(* IEC 61131-3 sources: daoli-st-library/DL_MathData (part 29) *)

(* ---- FB_DL_MovingAverage.st ---- *)
(*==============================================================================
 * 组件名称 (Component)  : FB_DL_MovingAverage
 * 所属子库 (Sublibrary) : DL_MathData
 * 当前版本 (Version)    : 1.0.0
 * 兼容性   (Platform)   : CODESYS 3.5 / TwinCAT 3 / 汇川 InoProShop / Machine Expert
 *                         仅依赖 Standard.library（R_TRIG），全 REAL 运算
 * 功能描述 (Function)   : O(1) 递推滑动平均滤波。窗口长度运行时可改，采样节拍由
 *                         调用方控制。两阶段启动：窗口未满阶段只"写入+累加+计数"、
 *                         绝不执行"减最旧值"；窗口已满阶段执行"减最旧+加最新+指针递增"。
 *                         每 DL_MAV_CORRECT_CYCLE 次采样做一次全窗口重算，消除浮点
 *                         累加漂移。窗口长度变更时整体重建缓冲区，避免新旧样本混算产生台阶。
 *
 * 【滞后披露 / Phase lag disclosure（边界 B11）】
 *   相位滞后约 (N-1)/2 个采样周期，滤波时间窗 = N × 采样周期。
 *   安全联锁回路（急停、超压保护、超温切断）严禁使用大窗口滤波值，
 *   必须直接使用原始信号或小窗口（N ≤ 3）值。
 *
 * 【断电保持提示 / Retain hint（边界 B12）】
 *   缓冲区、写指针、累加和、已填充数若不设 RETAIN，重新上电会重走"窗口未满"阶段，
 *   表现为输出从 0 缓慢爬升。需要无扰重启的场合，应将本实例声明为 VAR RETAIN。
 *
 * 【采样语义 / Sampling semantics（边界 B7，重要）】
 *   采样判据统一为"bSample 电平为 TRUE 即采样"：bSample := TRUE 常 TRUE 时每周期采样，
 *   接一个上升沿脉冲变量则按事件采样。绝不用 R_TRIG 承担两种语义——常 TRUE 信号经
 *   R_TRIG 只在首周期产生一次脉冲，会导致"只采到一个样本"的低级事故。
 *   因此本组件不设 fbTrigSample 采样沿实例（仅保留 fbTrigReset），
 *   这是对 ROUND_PLAN §2.13 VAR 清单的刻意收窄，依据 B7 与决策记录 P6。
 *
 * 【状态机 / State machine（边界 B1/B10）】
 *   采用 eInit / eFilling / eRunning / eFault 四态 + ELSE 兜底。
 *   两阶段判据由 bBufferFull 承担并在采样段用 IF bBufferFull THEN … ELSE … END_IF（代码骨架，示例省略）
 *   显式分支，采样算术只写一处，状态机只负责阶段迁移，避免同一段代码在两个 CASE
 *   分支中重复而导致"只改一处"的缺陷。
 * 开源溯源 (Origin)     : 原创实现。环形缓冲 + 递推求和的滑动平均为公开经典算法。
 * 依赖     (Depends)    : 无 DL_ 内部依赖；Standard.library: R_TRIG
 * 红线自检 (Redline)    : R1 ✓ 零全局变量表与外部变量引用 ｜ R2 ✓ 零物理 IO 地址直写
 *                         R3 ✓ 纯 IEC 61131-3 ｜ R4 ✓ 除零双保险/窗口钳位/MOD 回绕/重算防死锁
 *                         R5 ✓ 全变量中英双语同行注释 ｜ R6 ✓ 四态 ENUM+CASE+ELSE 兜底
 *                         R7 ✓ R_TRIG 主体最前部无条件刷新
 * 修订历史 (Revision)   :
 *   2026-11-14  v1.0.0  首版入库（Phase 1 冷启动 · Level 0 批次）
 *============================================================================*)

(*-----------------------------------------------------------------------------
 * 枚举: E_DL_MovingAverageState（归属 DL_MathData，与 FB_DL_MovingAverage 同文件）
 * 含义: 滑动平均工作阶段。eFilling 与 eRunning 的区分仅用于状态迁移与诊断，
 *       采样算术由 bBufferFull 在单一分支内完成。
 *----------------------------------------------------------------------------*)
TYPE E_DL_MovingAverageState :
(
    eInit    := 0,    // 初始化态：清缓冲、清累加和、清故障，单周期驻留 / Initialization: clear buffer, sum and fault, single scan
    eFilling := 10,   // 填充态：窗口未满，只追加样本不做淘汰 / Filling: window not full, append only without eviction
    eRunning := 20,   // 运行态：窗口已满，执行 O(1) 递推替换 / Running: window full, O(1) recursive replacement
    eFault   := 99    // 故障态：非法状态命中，输出保持最后有效值 / Fault: illegal state hit, outputs hold the last valid value
);
END_TYPE

FUNCTION_BLOCK FB_DL_MovingAverage
VAR_INPUT
    fInput      : REAL := 0.0;      // 原始采样值 [EU] / Raw sampled value [EU]
    nWindowSize : INT := 8;         // 窗口长度，合法域 1..100 / Window length, valid range 1..100
    bSample     : BOOL := TRUE;     // 采样触发，电平 TRUE 即采样；接脉冲变量则按事件采样 / Sample trigger, TRUE level samples every scan
    bEnable     : BOOL := TRUE;     // 使能标志，FALSE 时停止采样并保持输出 / Enable flag, FALSE stops sampling and holds the output
    bReset      : BOOL;             // 复位信号，上升沿清空窗口与累加和 / Reset, rising edge clears the buffer and the sum
END_VAR
VAR_OUTPUT
    fAverage     : REAL;            // 窗口算术平均 [EU] / Window arithmetic mean [EU]
    bBufferFull  : BOOL;            // 窗口已填满标志，同时作为两阶段判据 / Buffer full flag, also the two-phase discriminator
    nSampleCount : INT;             // 窗口内有效样本数，值域 0..nWindowSize / Valid sample count in the window, range 0..nWindowSize
    fWindowSum   : REAL;            // 窗口累加和，诊断用 [EU] / Window sum for diagnostics [EU]
    bError       : BOOL;            // 故障标志，需 bReset 清除 / Fault flag, cleared by bReset
    uErrorId     : UDINT;           // 故障码，0 = 无故障 / Error code, 0 = no error
END_VAR
VAR
    afBuffer     : ARRAY[0..99] OF REAL;  // 环形缓冲区，容量等于窗口上限 [EU] / Ring buffer sized to the max window [EU]
    nWriteIndex  : INT;             // 环形写指针，值域 0..99 / Ring write index, range 0..99
    nFilled      : INT;             // 已填充样本数，值域 0..100 / Number of filled samples, range 0..100
    fSum         : REAL;            // 滑动累加和 [EU]，与 nFilled 同步维护 / Running sum [EU], maintained with nFilled
    nLastWindow  : INT;             // 上周期窗口长度，用于变更检测 / Previous window length for change detection
    fbTrigReset  : R_TRIG;          // 复位上升沿检测实例 / Reset rising edge detector instance
    nCorrectCnt  : DINT;            // 距下次全窗口重算的采样计数 / Sample counter until the next full-window recalculation
    nGuard       : DINT;            // 重算循环防死锁计数器 / Recalculation loop deadlock guard
    fRecalcSum   : REAL;            // 重算中间累加和 [EU] / Recalculation intermediate sum [EU]
    nIdx         : INT;             // 重算循环索引，值域 0..99 / Recalculation loop index, range 0..99
    nWindowEff   : INT;             // 钳位后的有效窗口长度 / Clamped effective window length
    eState       : E_DL_MovingAverageState; // 主状态机当前状态 / Current state of the main state machine
    bDoSample    : BOOL;            // 本周期采样使能（bSample AND bEnable） / Sampling enabled this scan
    bJustReset   : BOOL;            // 本周期刚发生复位/初始化，需跳过采样 / Reset or init happened this scan, sampling is skipped
END_VAR
VAR CONSTANT
    DL_MAV_MAX_WINDOW    : INT := 100;        // 窗口上限，必须与数组维度一致 / Max window, must match the array dimension
    DL_MAV_MIN_WINDOW    : INT := 1;          // 窗口下限 / Min window
    DL_MAV_CORRECT_CYCLE : DINT := 10000;     // 每 N 次采样做一次全窗口重算校正 / Recalculate every N samples
    DL_MAV_MAX_LOOP      : DINT := 100;       // 重算循环迭代上限 / Recalculation loop iteration limit
    DL_FLOAT_EPS         : REAL := 1.0E-6;    // 浮点判零容差 / Float zero tolerance
END_VAR

(*------------------------------------------------------------------------------
 * 段 1｜无条件刷新区（红线 R7）：复位沿实例在主体最前部调用，严禁进入 IF/CASE
 *      Unconditional refresh zone: the reset edge instance runs at the very top
 *-----------------------------------------------------------------------------*)
fbTrigReset(CLK := bReset);

(*------------------------------------------------------------------------------
 * 段 2｜窗口长度钳位（边界 B3）：先钳位，后用于所有后续计算
 *      Window length clamping: clamp first, then use everywhere
 *------------------------------------------------------------------------------*)
IF nWindowSize < DL_MAV_MIN_WINDOW THEN
    nWindowEff := DL_MAV_MIN_WINDOW;
    uErrorId   := 16#0001_0001;
    bError     := TRUE;
ELSIF nWindowSize > DL_MAV_MAX_WINDOW THEN
    nWindowEff := DL_MAV_MAX_WINDOW;
    uErrorId   := 16#0001_0001;
    bError     := TRUE;
ELSE
    nWindowEff := nWindowSize;
END_IF

(*------------------------------------------------------------------------------
 * 段 3｜窗口长度变更重建（边界 B4）：清空缓冲、指针、累加和，重走未满阶段
 *      Window change rebuild: clear buffer, pointer and sum, restart the filling phase
 *      不清空会让新旧窗口样本混算，输出出现台阶，现场会误判为传感器跳变
 *-----------------------------------------------------------------------------*)
bJustReset := FALSE;

IF nWindowEff <> nLastWindow THEN
    nLastWindow  := nWindowEff;
    nWriteIndex  := 0;
    nFilled      := 0;
    fSum         := 0.0;
    nCorrectCnt  := 0;
    bBufferFull  := FALSE;
    eState       := eInit;
    bJustReset   := TRUE;
END_IF

(*------------------------------------------------------------------------------
 * 段 4｜复位处理（边界 B9）：复位优先于采样，本周期不再采样
 *      Reset handling: reset wins over sampling, no sample is taken this scan
 *-----------------------------------------------------------------------------*)
IF fbTrigReset.Q THEN
    eState      := eInit;
    bJustReset  := TRUE;
END_IF

(*------------------------------------------------------------------------------
 * 段 5｜主状态机（红线 R6 / 边界 B10）：四态迁移，ELSE 兜底进故障
 *      Main state machine: four-state transition with an ELSE fallback
 *------------------------------------------------------------------------------*)
CASE eState OF

    eInit:
        (* 清空全部累积量，进入填充阶段；故障与错误码同时清除（边界 B9） *)
        (* Clear all accumulators and enter filling; fault and error code are cleared too *)
        nWriteIndex := 0;
        nFilled     := 0;
        fSum        := 0.0;
        fAverage    := 0.0;
        fWindowSum  := 0.0;
        bBufferFull := FALSE;
        nCorrectCnt := 0;
        uErrorId    := 16#0000_0000;
        bError      := FALSE;
        eState      := eFilling;

    eFilling:
        (* 未满阶段：窗口填满即迁移到运行阶段 *)
        (* Filling phase: migrate to running once the window is full *)
        IF bBufferFull THEN
            eState := eRunning;
        END_IF

    eRunning:
        (* 满窗阶段：若窗口被放大导致已填样本不足，回退到填充阶段（边界 B4 配套） *)
        (* Running phase: fall back to filling if the window grew beyond the filled count *)
        IF NOT bBufferFull THEN
            eState := eFilling;
        END_IF

    eFault:
        (* 故障态：不采样、不清缓冲；锁存故障标志，输出由段 8 按最后有效累加值刷新 *)
        (* Fault state: no sampling, no buffer clearing; latch the fault flag, stage 8 holds the output *)
        bError := TRUE;

    ELSE
        (* 非法状态拦截：进入故障态并上报，不做隐式恢复 *)
        (* Illegal state interception: enter fault and report, no implicit recovery *)
        eState   := eFault;
        uErrorId := 16#0001_0005;
        bError   := TRUE;

END_CASE;

(*------------------------------------------------------------------------------
 * 段 6｜采样触发判定（边界 B8）：电平语义 + 使能串接，复位当周期不采样
 *      Sampling decision: level semantics AND enable, suppressed on a reset scan
 *-----------------------------------------------------------------------------*)
bDoSample := bSample AND bEnable AND NOT bJustReset AND (eState <> eFault);

(*------------------------------------------------------------------------------
 * 段 7｜采样与递推（边界 B1/B2/B5/B6，本组件核心）
 *      Sampling and recursion, the core of this block
 *-----------------------------------------------------------------------------*)
IF bDoSample THEN

    (* 写指针上下界双检（红线 R4）：MOD 已保证范围内，仍显式兜底防越界写 *)
    (* Write index double check: MOD already guarantees the range, kept as an explicit guard *)
    IF (nWriteIndex < 0) OR (nWriteIndex > (DL_MAV_MAX_WINDOW - 1)) THEN
        nWriteIndex := 0;
        uErrorId    := 16#0001_0001;
        bError      := TRUE;
    END_IF

    IF bBufferFull THEN
        (*----------------------------------------------------------------------
         * 段 7a｜窗口已满：O(1) 递推——减去写指针处的最旧样本，再写入最新样本
         *       Buffer full: O(1) recursion, subtract the oldest then write the newest
         *       满窗时写指针恰好指向最旧样本，一个指针同时承担写入位与淘汰位
         *---------------------------------------------------------------------*)
        fSum := fSum - afBuffer[nWriteIndex] + fInput;
        afBuffer[nWriteIndex] := fInput;
    ELSE
        (*----------------------------------------------------------------------
         * 段 7b｜窗口未满：只追加样本与累加，绝不执行"减最旧值"
         *       Buffer not full: append only, never subtract the oldest
         *       若此处也减最旧值，会减掉尚未写入的 0，输出被系统性压低，
         *       表现为上电初期滤波值比原始信号更抖——即经典的两阶段缺陷
         *---------------------------------------------------------------------*)
        afBuffer[nWriteIndex] := fInput;
        fSum      := fSum + fInput;
        nFilled   := nFilled + 1;

        IF nFilled >= nWindowEff THEN
            nFilled     := nWindowEff;
            bBufferFull := TRUE;
        END_IF
    END_IF

    (*--------------------------------------------------------------------------
     * 段 7c｜指针回绕（边界 B5）：必须用 MOD，除数已由段 2 保证 ≥ 1
     *       Pointer wrap: MOD is mandatory, the divisor is guaranteed ≥ 1 by stage 2
     *-------------------------------------------------------------------------*)
    nWriteIndex := (nWriteIndex + 1) MOD nWindowEff;

    (*--------------------------------------------------------------------------
     * 段 7d｜浮点累加漂移校正（边界 B6）：每 N 次采样做一次全窗口重算
     *       Drift correction: a full-window recalculation every N samples
     *       FOR 循环设迭代上限并 EXIT，防止异常数据把扫描周期拖死
     *-------------------------------------------------------------------------*)
    nCorrectCnt := nCorrectCnt + 1;

    IF nCorrectCnt >= DL_MAV_CORRECT_CYCLE THEN
        nCorrectCnt := 0;
        fRecalcSum  := 0.0;
        nGuard      := 0;

        FOR nIdx := 0 TO (nFilled - 1) DO
            IF (nIdx >= 0) AND (nIdx <= (DL_MAV_MAX_WINDOW - 1)) THEN
                fRecalcSum := fRecalcSum + afBuffer[nIdx];
            END_IF

            nGuard := nGuard + 1;

            IF nGuard >= DL_MAV_MAX_LOOP THEN
                EXIT;
            END_IF
        END_FOR;

        fSum := fRecalcSum;
    END_IF

END_IF

(*------------------------------------------------------------------------------
 * 段 8｜输出刷新（边界 B2）：除零双保险——窗口钳位已保证 nWindowEff ≥ 1，
 *      此处再以 nFilled > 0 兜底，两道防线缺一不可
 *      Output refresh: dual divide-by-zero protection, both guards are mandatory
 *      使能关闭时 nFilled 与 fSum 不变，平均值自然保持，不清空缓冲区（边界 B8）
 *-----------------------------------------------------------------------------*)
fWindowSum   := fSum;
nSampleCount := nFilled;

IF nFilled > 0 THEN
    fAverage := fSum / INT_TO_REAL(nFilled);
ELSE
    fAverage := 0.0;
END_IF
END_FUNCTION_BLOCK

(* ---- FB_DL_RingBufferLReal.st ---- *)
(*==============================================================================
 * 组件名称 (Component)  : FB_DL_RingBufferLReal
 * 所属子库 (Sublibrary) : DL_MathData
 * 当前版本 (Version)    : 1.0.0
 * 兼容性   (Platform)   : CODESYS 3.5 / TwinCAT 3 / 汇川 InoProShop / Machine Expert
 *                         仅依赖 Standard.library（R_TRIG），浮点用标准 64 位类型
 * 功能描述 (Function)   : 定长 64 容量的 LREAL 环形队列（先进先出）。压入 / 弹出 / 窥视 /
 *                         清空四操作全部 O(1)，无任何元素搬移与循环。
 *                         解决"每来一个样本把整段数组移位一次还容易错位一格"、
 *                         "故障前最后一段数据被冲掉无法追溯"两类现场问题。
 *                         满时拒绝写入而不覆盖最旧值：FIFO 语义下静默覆盖会让
 *                         数据丢失变得不可见，需要滑动窗口语义的场合请用滑动平均块。
 *                         全部指针更新只用"加一后取模"的前向回绕，
 *                         组件内不存在任何指针减法，从结构上规避负数取模的平台差异。
 * 开源溯源 (Origin)     : 原创实现。环形队列 + 计数区分空满为公开经典算法；
 *                         本库仅借鉴其 O(1) 递推语义，独立重构，未复制任何源码。
 * 本文件内含       : FB    FB_DL_RingBufferLReal（单 POU，无配套类型）
 * 依赖     (Depends)    : 无 DL_ 内部依赖；Standard.library: R_TRIG
 * 红线自检 (Redline)    : R1 ✓ 禁用全局存储与物理寻址 ｜ R2 ✓ 无地址直写
 *                         R3 ✓ 纯 IEC 61131-3，计数比较显式转换 ｜ R4 ✓ 下标双检 + 前向取模回绕
 *                         R5 ✓ 全变量中英双语同行注释 ｜ R6 N/A（队列无跨周期状态转移，指针与计数即全部状态）
 *                         R7 ✓ 两 R_TRIG 主体最前部无条件刷新 ｜ R8 ✓ 容量常量化
 *
 * 【容量与内存披露 / Capacity and memory（边界 B10）】
 *   固定容量 64 元素，元素为 64 位浮点，实例净占用约 512 字节缓冲区，
 *   加指针与计数共约 0.6KB。定长数组跨平台行为一致，运行时容量参数化
 *   会引入动态数组差异，故不提供。
 *
 * 【哨兵值披露 / Sentinel disclosure（边界 B7）】
 *   空队时窥视输出 0.0，该 0.0 是哨兵不是数据。判空必须看空标志，
 *   不得以"窥视值等于 0"反推队列状态——0 是合法的采样值。
 *
 * 【同周期压弹次序 / Push-before-pop ordering（边界 B5）】
 *   同一扫描周期同时出现压入沿与弹出沿时，先压后弹，净效果为"换出队首"。
 *   该次序不可交换，改动会改变满队与单元素队列的行为语义。
 *
 * 修订历史 (Revision)   :
 *   2026-11-14  v1.0.0  首版入库（Phase 1 第二轮 · Level 0 批次 C）
 *============================================================================*)
FUNCTION_BLOCK FB_DL_RingBufferLReal
VAR_INPUT
    fPushValue : LREAL;   // 待压入值 [EU] / Value to push [EU]
    bPush      : BOOL;    // 上升沿压入 / Push on rising edge
    bPop       : BOOL;    // 上升沿弹出 / Pop on rising edge
    bClear     : BOOL;    // 电平清空，最高优先级操作 / Level-triggered clear, highest priority
END_VAR
VAR_OUTPUT
    fPopValue  : LREAL;   // 最近一次弹出值 [EU]，空读被拒时保持上次值 / Last popped value [EU], holds on a rejected pop
    fPeekValue : LREAL;   // 队首值 [EU]，空队时为 0.0 哨兵 / Front value [EU], 0.0 sentinel when empty
    uCount     : UINT;    // 当前元素数 [个]，值域 0..64 / Current element count [count], range 0..64
    bFull      : BOOL;    // 已满标志 / Full flag
    bEmpty     : BOOL;    // 已空标志 / Empty flag
    uErrorId   : UDINT;   // 故障码，0 = 无故障 / Error code, 0 = no error
END_VAR
VAR
    afBuffer   : ARRAY[0..63] OF LREAL;  // 环形存储区 [EU] / Ring storage [EU]
    nReadIdx   : INT;                    // 读指针（队首），值域 0..63 / Read index (front), range 0..63
    nWriteIdx  : INT;                    // 写指针（下一写入位），值域 0..63 / Write index (next slot), range 0..63
    fbTrigPush : R_TRIG;                 // 压入沿检测实例 / Push edge detector instance
    fbTrigPop  : R_TRIG;                 // 弹出沿检测实例 / Pop edge detector instance
END_VAR
VAR CONSTANT
    DL_RB_CAP : INT := 64;   // 固定容量，必须与数组维度严格一致 / Fixed capacity, must match the array
END_VAR

(*------------------------------------------------------------------------------
 * 段 1｜无条件刷新区（红线 R7）：两个边沿实例位于主体最前部，严禁进入 IF / CASE
 *      Unconditional refresh zone: both edge instances run at the very top
 *-----------------------------------------------------------------------------*)
fbTrigPush(CLK := bPush);
fbTrigPop(CLK  := bPop);

(*------------------------------------------------------------------------------
 * 段 2｜故障码本周期清零
 *      Error code is cleared every scan
 *-----------------------------------------------------------------------------*)
uErrorId := 16#0000_0000;

(*------------------------------------------------------------------------------
 * 段 3｜清空（边界 B2）：电平触发、最高优先级，先于压弹处理
 *      Clear: level-triggered and highest priority, handled before push and pop
 *      这样"清空与压入同周期"的结果只可能是"压入一个元素"，不存在歧义
 *      Clear-then-push in one scan deterministically leaves exactly one element
 *-----------------------------------------------------------------------------*)
IF bClear THEN
    nReadIdx  := 0;
    nWriteIdx := 0;
    uCount    := UINT#0;
    fPeekValue := 0.0;
ELSE

    (*--------------------------------------------------------------------------
     * 段 4｜压入（边界 B3）：满时拒绝写入，绝不覆盖最旧值
     *      Push: rejected when full, the oldest value is never silently overwritten
     *-------------------------------------------------------------------------*)
    IF fbTrigPush.Q THEN
        IF uCount >= INT_TO_UINT(DL_RB_CAP) THEN
            uErrorId := 16#0001_0009;
        ELSE
            (* 写指针双检：MOD 已保证范围，仍显式兜底防越界写（R4） *)
            (* Write index double check, kept as an explicit guard besides MOD *)
            IF (nWriteIdx >= 0) AND (nWriteIdx < DL_RB_CAP) THEN
                afBuffer[nWriteIdx] := fPushValue;
            ELSE
                nWriteIdx := 0;
                afBuffer[nWriteIdx] := fPushValue;
            END_IF

            (* 前向取模回绕：组件内不存在指针减法（边界 B6） *)
            (* Forward modulo wrap, no pointer subtraction anywhere in this component *)
            nWriteIdx := (nWriteIdx + 1) MOD DL_RB_CAP;
            uCount    := uCount + UINT#1;
        END_IF
    END_IF

    (*--------------------------------------------------------------------------
     * 段 5｜弹出（边界 B4/B5）：空时拒绝，弹出值保持上次有效值
     *      Pop: rejected when empty, the last valid value is held
     *      与压入同周期出现时按"先压后弹"处理，此处已位于压入之后
     *      Handled after the push stage, implementing the push-before-pop order
     *-------------------------------------------------------------------------*)
    IF fbTrigPop.Q THEN
        IF uCount = UINT#0 THEN
            uErrorId := 16#0001_000A;
        ELSE
            IF (nReadIdx >= 0) AND (nReadIdx < DL_RB_CAP) THEN
                fPopValue := afBuffer[nReadIdx];
            ELSE
                nReadIdx  := 0;
                fPopValue := afBuffer[nReadIdx];
            END_IF

            nReadIdx := (nReadIdx + 1) MOD DL_RB_CAP;
            uCount   := uCount - UINT#1;
        END_IF
    END_IF

    (*--------------------------------------------------------------------------
     * 段 6｜窥视（边界 B7）：每周期刷新队首，空队输出哨兵 0.0
     *      Peek: refreshed every scan, the empty queue reports the 0.0 sentinel
     *-------------------------------------------------------------------------*)
    IF uCount > UINT#0 THEN
        IF (nReadIdx >= 0) AND (nReadIdx < DL_RB_CAP) THEN
            fPeekValue := afBuffer[nReadIdx];
        ELSE
            fPeekValue := 0.0;
        END_IF
    ELSE
        fPeekValue := 0.0;
    END_IF

END_IF

(*------------------------------------------------------------------------------
 * 段 7｜状态标志（边界 B8）：空满由计数派生，计数只在成功路径上加减
 *      Status flags: derived from the count, which only moves on success paths
 *-----------------------------------------------------------------------------*)
bFull  := (uCount >= INT_TO_UINT(DL_RB_CAP));
bEmpty := (uCount = UINT#0);
END_FUNCTION_BLOCK

(* ---- FB_DL_ScaleRangeWatch.st ---- *)
(*
    FB_DL_ScaleRangeWatch —— 工程量标定区间越界监视（回差 + 延时确认 + 故障锁存）
    ------------------------------------------------------------------
    组件名称  : FB_DL_ScaleRangeWatch
    分类      : DL_MathData / Scaling
    前缀      : FB_DL_
    版本      : 1.0.1
    溯源      : 借鉴点 —— 过程仪表标定链的通行三段式：原始码 → 工程量线性换算
                → 带迟滞与延时确认的上下限越界判定；该「换算 + 越界监测」组合
                在开源数学/测量库族中属常见语义，本件借鉴其**判据顺序与迟滞口径**，
                不借用其任何数据结构、命名或代码组织。
                clean-room 声明 —— 零代码行复制；换算仅用标准运算符，定时与
                沿检测仅用 IEC 61131-3 标准库 TON / R_TRIG。
                许可证 —— 本件 MIT；来源标签 lgf-math 仅作语义参考，
                本件不包含、不派生其任何受版权保护的实现。
    平台      : 纯 IEC 61131-3，CODESYS 3.5 / TwinCAT 3 / InoProShop / Machine Expert 通用
    作者      : 道莅代码库 · PLC编程专家（R70 构建轮 · 批 1 · N3）
    ------------------------------------------------------------------
    功能说明  : fEng = fRaw * fGain + fOffset，随后对 fEng 判上下限：
                越过 fHighLim 且持续 tConfirm 才置 bHighAlarm，跌回
                fHighLim - fHyst 才复位；下限对称（fLowLim / fLowLim + fHyst）。
                定时器无条件周期调用（规则 ⑦），IN 用显式条件表达式，
                且条件中已把「已报警自保持」并入，故复位只由回差线决定，
                不存在无回差抖振。
                故障锁存口径（R187 / R189）：组态非法或原始值非有限 → 锁存首个
                成因码至 _nCodeLatch，bReset 上升沿解除；**故障期内不按当下输入
                重新推断成因**，一律回放锁存码，避免成因漂移。
                换算除法面：本件无除法（增益为乘子），无除零面；
                但增益为 0 属**增益零域**（v1.0.1 起拦截，见边界六）：
                fGain = 0.0 时 fEng ≡ fOffset，工程量被钉死在偏置值，
                上下限报警将永久不触发（保护静默失效），故按组态非法处理。
    错误码    : 16#0002_0121 组态非法（v1.0.1 起含增益零域成因），锁存，输出清零 —— 故障级
                16#0002_0122 原始值非有限，锁存，输出保持末次良好工程值 —— 故障级
    码位总账  : 16#0002_0121 用 ｜ 16#0002_0122 用
    状态机    : N/A —— 单相监视，无顺序状态机，无 ENUM / CASE 可写；
                两路确认计时由 TON 实例自持，属定时器状态而非顺序状态
    边界与披露: 一 组态判据逐项点名（R272）：fGain / fOffset / fHighLim / fLowLim /
                   fHyst 全部纳入非有限闸；fHighLim <= fLowLim 拦截；fHyst < 0 拦截；
                   fHyst >= (fHighLim - fLowLim) 拦截（迟滞吞没整带时上下限无回差带，
                   判据恒真）；tConfirm < T#0S 不可表示，故不设该判据；
                二 输入非有限时 fEng 输出**保持末次良好值**（_bHaveGood 为真才输出，
                   否则输出 0.0），并在头注释声明该保持语义（R191 名实双出口）；
                三 失能（bEn = FALSE）语义写死（R303）：fEng 输出 0.0、bHighAlarm /
                   bLowAlarm / bInBand / bBusy 全清零、nErrCode 清零、bError 清零，
                   但 _bFault 锁存位**不被失能清除**（失能是操作态，不是复位），
                   必须 bReset 上升沿才解除 —— 两者语义分离，避免失能顺手清故障；
                四 定时器 _tonHigh / _tonLow 无论失能 / 故障 / 正常均在段 9 无条件调用，
                   IN 为段 8 计算出的显式条件，未放入任何可能被跳过的分支；
                五 量程零域拦截路径（v1.0.1 点修，缺陷 H4）：fGain = 0.0（增益零域，
                   判据 ABS(fGain) <= DL_SRW_GMIN，GMIN = 1.0E-15）时 fEng ≡ fOffset，
                   工程量被钉死在偏置值，上下限报警永久不触发且无任何故障码 ——
                   保护静默失效，比除零更隐蔽；v1.0.1 起段 4 组态闸并联该判据，
                   增益零域 → 码 0121 组态锁存、段 8 换算段结构性不可达、报警不静默；
                六 零域第二道判据（v1.0.0 既有，H2 复核确认）：fHighLim <= fLowLim
                   对 fHighLim = fLowLim 的零带宽路径同样拦截，两道判据冗余覆盖
                   零量程，不存在可进入段 8 换算段的零域反例向量（±1E30 极端
                   幅值下带宽差 <= 2E30 < LREAL 域，无溢出面）；
                七 复位解除当拍语义（H3 披露，行为不变）：段 3 清锁存与段 6 同拍
                   重判组态发生在同一扫描周期，组态仍非法则同拍重锁存 —— 与
                   R189 口径一致，非缺陷，仅声明；
                八 段 8 非有限换算分支就地锁存 0121，不含「增益 × 原始值溢出」
                   独立成因项 —— 溢出归因为组态域外（增益超域），与 R190 归因
                   唯一口径不冲突，声明即可；
                九 零全局变量、零 VAR_EXTERNAL、零物理地址、零数组下标。
    修订记录  : 2026-11-22 v1.0.0 首次入库（R70 构建轮 · 批 1 · N3）
                2026-11-22 v1.0.1 点修（R71 · 批 1 · 序号 1）：段 4 组态闸并联
                增益零域判据 ABS(fGain) <= DL_SRW_GMIN（缺陷 H4，R70 挂账复核），
                新增常量 DL_SRW_GMIN = 1.0E-15；码位沿用 16#0002_0121 不新开；
                头注释补量程零域拦截路径披露与复位当拍重锁存语义声明；
                不改引脚、不改其他段行为（H1 文档-源码口径漂移已以源码实测对账）。
*)
FUNCTION_BLOCK FB_DL_ScaleRangeWatch
VAR_INPUT
    fRaw      : LREAL;                     (* 原始值（未标定，可为 ADC 码或物理量），[原始单位] / the raw unscaled value *)
    fGain     : LREAL := 1.0;              (* 标定增益（斜率），[工程单位/原始单位] / the calibration gain, the slope *)
    fOffset   : LREAL := 0.0;              (* 标定偏置（截距），[工程单位] / the calibration offset, the intercept *)
    fHighLim  : LREAL := 100.0;            (* 上限判据值，[工程单位]，须 > fLowLim / the upper limit, must exceed fLowLim *)
    fLowLim   : LREAL := 0.0;              (* 下限判据值，[工程单位]，须 < fHighLim / the lower limit, must be under fHighLim *)
    fHyst     : LREAL := 0.0;              (* 回差带宽，[工程单位]，域 [0, fHighLim - fLowLim) / the hysteresis band *)
    tConfirm  : TIME := T#1S;              (* 越界确认延时，[ms]，须 >= T#0S / the out-of-range confirmation delay *)
    bEn       : BOOL := TRUE;              (* 使能，[标志]，FALSE 时出口清零（R303）/ the enable, FALSE clears the outlets *)
    bReset    : BOOL := FALSE;             (* 故障复位，[标志]，上升沿解除锁存 / the reset, its rising edge clears the latch *)
END_VAR
VAR_OUTPUT
    fEng      : LREAL;                     (* 换算后工程值，[工程单位] / the scaled engineering value *)
    bHighAlarm : BOOL;                     (* 上限越界报警（回差 + 延时确认后），[标志] / the high limit alarm *)
    bLowAlarm : BOOL;                      (* 下限越界报警（回差 + 延时确认后），[标志] / the low limit alarm *)
    bInBand   : BOOL;                      (* 工程值在带内（两侧报警均为假），[标志] / the value sits inside the band *)
    bBusy     : BOOL;                      (* 确认计时进行中（越界已出现但未满延时），[标志] / a confirmation timer is running *)
    bValid    : BOOL;                      (* 输出可用，故障或失能为 FALSE / the outlets are usable *)
    bError    : BOOL;                      (* 故障标志，存在锁存故障时为 TRUE / the fault flag, raised on a latched fault *)
    nErrCode  : UDINT;                     (* 错误码，0 = 正常，锁存回放 / the error id, 0 = ok, replayed from the latch *)
END_VAR
VAR
    _rtReset   : R_TRIG;                   (* 复位上升沿检测实例（无条件调用）/ the reset rising edge instance *)
    _tonHigh   : TON;                      (* 上限确认延时实例（无条件调用）/ the high limit confirmation timer *)
    _tonLow    : TON;                      (* 下限确认延时实例（无条件调用）/ the low limit confirmation timer *)
    _bFault    : BOOL;                     (* 故障锁存位，仅 bReset 上升沿解除 / the latched fault bit *)
    _nCodeLatch : UDINT;                   (* 锁存成因码，故障期回放 / the latched cause code, replayed while faulted *)
    _bCfgBad   : BOOL;                     (* 组态非法标志（逐拍重算，仅用于首次锁存）/ the configuration fault flag *)
    _bInBad    : BOOL;                     (* 原始值非有限标志（逐拍重算，仅用于首次锁存）/ the input fault flag *)
    _bRun      : BOOL;                     (* 运行许可 = 使能 且 无锁存故障 / the run permit *)
    _bHighCond : BOOL;                     (* 上限确认条件（含自保持与回差，送 TON）/ the high confirmation condition *)
    _bLowCond  : BOOL;                     (* 下限确认条件（含自保持与回差，送 TON）/ the low confirmation condition *)
    _fEngTmp   : LREAL;                    (* 换算中间量，[工程单位] / the scaling temporary *)
    _fLastGood : LREAL;                    (* 末次良好工程值，[工程单位] / the last good engineering value *)
    _bHaveGood : BOOL;                     (* 已获得过良好值，[标志] / a good value has been seen *)
END_VAR
VAR CONSTANT
    DL_SRW_FMAX : LREAL := 1.0E30;         (* 非有限筛查幅值上限，[工程单位] / the finiteness screening cap *)
    DL_SRW_GMIN : LREAL := 1.0E-15;        (* 增益零域判据阈值，|fGain| <= 此值视为零增益组态非法，[无量纲] / the zero-gain threshold, |fGain| <= this means an illegal zero-gain configuration *)
END_VAR

// 段 1｜出口预置（统一出口预置，R256）/ segment 1, preset every outlet
fEng       := 0.0;                         // 工程值预置 0.0 / preset the engineering value to zero
bHighAlarm := FALSE;                       // 上限报警预清零 / preset the high alarm false
bLowAlarm  := FALSE;                       // 下限报警预清零 / preset the low alarm false
bInBand    := FALSE;                       // 带内标志预清零 / preset the in-band flag false
bBusy      := FALSE;                       // 忙碌标志预清零 / preset the busy flag false
bValid     := FALSE;                       // 可用标志预清零 / preset the valid flag false
bError     := FALSE;                       // 故障标志预清零 / preset the error flag false
nErrCode   := 0;                           // 错误码预置无错 / preset the code to zero
_bHighCond := FALSE;                       // 上限条件预清零 / preset the high condition false
_bLowCond  := FALSE;                       // 下限条件预清零 / preset the low condition false

// 段 2｜复位沿检测（无条件调用，规则 ⑦）/ segment 2, the reset edge instance, called unconditionally
_rtReset(CLK := bReset);                   // 每周期无条件刷新 / refreshed every scan without exception

// 段 3｜锁存解除：仅 bReset 上升沿，锁存码同步清零 / segment 3, the latch release on the reset rising edge
IF _rtReset.Q THEN                         // 复位上升沿 / the reset rising edge
    _bFault     := FALSE;                  // 解除故障锁存 / release the fault latch
    _nCodeLatch := 0;                      // 清锁存码（可到达的清除边，R188）/ clear the latched code, a reachable clearing edge
END_IF

// 段 4｜组态守卫（边界一逐项点名 + 增益零域 H4，R272）/ segment 4, the configuration guard
_bCfgBad := (fHighLim <= fLowLim)                                        // 上下限反置或重合（兼拦零带宽，边界六）/ the limits reversed or coincident
         OR (fHyst < 0.0)                                                // 回差为负 / a negative hysteresis
         OR (fHyst >= (fHighLim - fLowLim))                              // 回差吞没整带 / the hysteresis swallows the band
         OR (ABS(fGain) <= DL_SRW_GMIN)                                  // 增益零域（H4，v1.0.1 起拦截）/ the zero-gain domain, intercepted since v1.0.1
         OR (fGain <> fGain) OR ((fGain - fGain) <> 0.0) OR (ABS(fGain) > DL_SRW_FMAX)        // 增益非有限 / the gain non finite
         OR (fOffset <> fOffset) OR ((fOffset - fOffset) <> 0.0) OR (ABS(fOffset) > DL_SRW_FMAX) // 偏置非有限 / the offset non finite
         OR (fHighLim <> fHighLim) OR ((fHighLim - fHighLim) <> 0.0) OR (ABS(fHighLim) > DL_SRW_FMAX) // 上限非有限 / the upper limit non finite
         OR (fLowLim <> fLowLim) OR ((fLowLim - fLowLim) <> 0.0) OR (ABS(fLowLim) > DL_SRW_FMAX)      // 下限非有限 / the lower limit non finite
         OR (fHyst <> fHyst) OR ((fHyst - fHyst) <> 0.0) OR (ABS(fHyst) > DL_SRW_FMAX);               // 回差非有限 / the hysteresis non finite

// 段 5｜输入守卫（NaN 自反判 + Inf 差值自反判 + 幅值上界）/ segment 5, the raw input guard
_bInBad := (fRaw <> fRaw) OR ((fRaw - fRaw) <> 0.0) OR (ABS(fRaw) > DL_SRW_FMAX); // 原始值非有限 / the raw value non finite

// 段 6｜首次成因锁存（故障期内不重推断，回放锁存码，R189）/ segment 6, the first-cause latch
IF NOT _bFault THEN                        // 未锁存时才有资格登记成因 / a cause is registered only while not latched
    IF _bCfgBad THEN                       // 组态非法（优先归因，组态是根因）/ an illegal configuration, the root cause first
        _bFault     := TRUE;               // 置故障锁存 / latch the fault
        _nCodeLatch := 16#0002_0121;       // 故障级：组态非法 / fault level: the configuration is illegal
    ELSIF _bInBad THEN                     // 原始值非有限 / the raw value is non finite
        _bFault     := TRUE;               // 置故障锁存 / latch the fault
        _nCodeLatch := 16#0002_0122;       // 故障级：输入非有限 / fault level: the input is non finite
    END_IF
END_IF

// 段 7｜运行许可：失能或锁存故障即退出换算 / segment 7, the run permit
_bRun := bEn AND NOT _bFault;              // 使能且无锁存故障 / enabled and not latched

// 段 8｜换算与条件计算（分支内不调用任何定时器）/ segment 8, the scaling and the conditions
IF _bRun THEN                              // 运行许可成立 / the run permit holds
    _fEngTmp := fRaw * fGain + fOffset;    // 工程量换算（委托 `*` 与 `+`）/ the engineering conversion, delegated
    IF (_fEngTmp <> _fEngTmp) OR ((_fEngTmp - _fEngTmp) <> 0.0) THEN // 换算结果非有限（增益超域导致）/ the result non finite
        _bFault     := TRUE;               // 就地锁存（增益巨大导致的溢出同属组态问题）/ latch in place
        _nCodeLatch := 16#0002_0121;       // 故障级：组态非法（增益域外）/ fault level: an illegal configuration
        fEng        := _fLastGood;         // 保持末次良好值（R191 名实双出口）/ hold the last good value
        bValid      := _bHaveGood;         // 有良好值才可用 / usable only if a good value was seen
        bError      := TRUE;               // 故障标志置位 / raise the fault flag
        nErrCode    := _nCodeLatch;        // 回放锁存码 / replay the latched code
    ELSE                                   // 换算结果有限 / the result is finite
        _fLastGood := _fEngTmp;            // 刷新末次良好值 / refresh the last good value
        _bHaveGood := TRUE;                // 标记已有良好值 / mark that a good value exists
        fEng       := _fEngTmp;            // 工程值出口 / the engineering outlet
        _bHighCond := (fEng > fHighLim) OR (_tonHigh.Q AND NOT (fEng < (fHighLim - fHyst))); // 上限条件：置位线或「已报警且未破回差线」
        _bLowCond  := (fEng < fLowLim) OR (_tonLow.Q AND NOT (fEng > (fLowLim + fHyst)));    // 下限条件：置位线或「已报警且未破回差线」
    END_IF
ELSE                                       // 失能或锁存故障 / disabled or latched
    bValid   := FALSE;                     // 输出不可用 / the outlets are unusable
    _bHighCond := FALSE;                   // 条件清零，计时器随之复位 / clear the condition, the timer resets
    _bLowCond  := FALSE;                   // 条件清零 / clear the condition
    IF NOT bEn THEN                        // 失能优先于故障归因（操作态，边界三）/ a disable takes precedence, an operator state
        fEng     := 0.0;                   // 失能相出口清零（R303）/ zero the outlet while disabled
        bError   := FALSE;                 // 失能不是故障 / a disabled block is not a fault
        nErrCode := 0;                     // 失能不发码 / no code while disabled
    ELSE                                   // 锁存故障相 / the latched fault phase
        fEng     := _fLastGood;            // 保持末次良好值（边界二，R191 名实双出口）/ hold the last good value
        bError   := _bFault;               // 故障位与锁存同源 / both outlets share the latch
        nErrCode := _nCodeLatch;           // 回放锁存码（不按当下输入重推断）/ replay the latched code
    END_IF
END_IF

// 段 9｜定时器无条件周期调用（规则 ⑦，IN 为显式条件）/ segment 9, unconditional timer calls
_tonHigh(IN := _bHighCond, PT := tConfirm);   // 上限确认计时，每周期无条件刷新 / the high confirmation timer
_tonLow(IN := _bLowCond, PT := tConfirm);     // 下限确认计时，每周期无条件刷新 / the low confirmation timer

// 段 10｜报警与忙碌出口（全部取自定时器 Q，单点写入）/ segment 10, the alarm and busy outlets
bHighAlarm := _bRun AND _tonHigh.Q;        // 上限报警：运行中且确认完成 / the high alarm, confirmed while running
bLowAlarm  := _bRun AND _tonLow.Q;         // 下限报警：运行中且确认完成 / the low alarm, confirmed while running
bInBand    := _bRun AND NOT bHighAlarm AND NOT bLowAlarm; // 带内：运行中且两侧均无报警 / inside the band
bBusy      := _bRun AND ((_bHighCond AND NOT _tonHigh.Q) OR (_bLowCond AND NOT _tonLow.Q)); // 确认计时进行中
IF _bRun AND _bHaveGood THEN               // 运行中且已有良好值 / running with a good value available
    bValid := TRUE;                        // 工程值可用 / the engineering value is usable
END_IF
END_FUNCTION_BLOCK

(* ---- FB_DL_ShrinkFilmUsageCalc.st ---- *)
(*
  Component : FB_DL_ShrinkFilmUsageCalc
  Category  : DL_MathData
  Type      : FB
  Version   : 1.0.0
  CodeSeg   : 16#02_3_5D
  Summary   : 收缩膜单包耗量换算与成本核算：膜长×膜宽×厚度→重量折算，按产量包数对齐口径出总耗与成本。
              Shrink film usage per pack and cost accounting: length x width x thickness to weight, aligned with pack count.
  溯源声明  : 道莅自研 clean-room
  边界安全  : 密度/厚度/膜长/膜宽正域闸（> 0，防除零与负值换算）；包数域闸（≥ 1，防产量口径为 0 除零）；
              价格非负域闸（≥ 0）；厚度 um→m 显式 1.0E-6 换算链，密度 g/cm³→kg/m³ ×1000；
              累计计数防 UDINT 回卷；全浮点比较带 fEps 容差。
  复用      : 无
*)

FUNCTION_BLOCK FB_DL_ShrinkFilmUsageCalc
VAR_INPUT
    bRun         : BOOL;               (* 核算使能，假则输出冻结 · Enable, FALSE freezes outputs *)
    fFilmLenM    : LREAL;              (* 单包膜长 [m] · Film length per pack *)
    fFilmWidthM  : LREAL;              (* 膜宽 [m] · Film width *)
    fThickUm     : LREAL;              (* 膜厚 [um] · Film thickness *)
    fDensityGcc  : LREAL := 0.92;      (* 膜密度 [g/cm³] · Film density *)
    fPriceYuanKg : LREAL := 12.0;      (* 膜价 [元/kg] · Film price *)
    nPackCnt     : INT;                (* 产量包数 [包]，口径对齐基准 · Production pack count *)
    fEps         : LREAL := 1.0E-6;    (* 浮点判零容差 [实数域] · Floating zero tolerance *)
END_VAR
VAR_OUTPUT
    fPerPackKg     : LREAL;            (* 单包耗膜重量 [kg] · Film weight per pack *)
    fTotalKg       : LREAL;            (* 总耗膜重量 [kg]（产量口径）· Total film weight *)
    fCostYuan      : LREAL;            (* 总成本 [元] · Total cost *)
    fCostPerPackYn : LREAL;            (* 单包成本 [元/包] · Cost per pack *)
    fTotalKgAcc    : LREAL;            (* 累计耗膜重量 [kg]，班次台账 · Cumulative weight ledger *)
    fCostYuanAcc   : LREAL;            (* 累计成本 [元]，班次台账 · Cumulative cost ledger *)
    bLedgerClr     : BOOL;             (* 台账清零指令 [事件]，真则清累计 · Ledger clear command *)
    bError         : BOOL;             (* 故障标志，与故障码配对 · Fault flag paired with codes *)
    uErrorId       : UDINT;            (* 事件码 16#0000_005D，0 无事件 · Event code *)
END_VAR
VAR
    uCode   : WORD;     (* 码位暂存，每拍重算 [码] · Code staging, recomputed *)
    bDimOk  : BOOL;     (* 尺寸域有效标志 · Dimension validity flag *)
    bCntOk  : BOOL;     (* 包数/价格域有效标志 · Count and price validity flag *)
    fDenGcc3: LREAL;    (* 密度 SI 换算值 [kg/m³] · Density in SI units *)
    fThickM : LREAL;    (* 厚度 SI 换算值 [m] · Thickness in SI units *)
    nCycles : UDINT;    (* 有效核算拍计数 [拍]，防回卷 · Valid calculation count with wrap guard *)
END_VAR
VAR CONSTANT
    DL_SFC_UM2M  : LREAL := 1.0E-6;    (* um 到 m 系数 [m/um] · Micrometers to meters *)
    DL_SFC_G2KG  : LREAL := 1000.0;    (* g/cm³ 到 kg/m³ 系数 · Gram per cc to kg per m3 *)
    DL_SFC_WRAP  : UDINT := 4294967290; (* 计数防回卷余量 [拍] · Counter wrap guard *)
END_VAR

(* === 段 0 · 实例刷新 === *)
(* 纯核算件：无 TON/R_TRIG 实例，计数状态见段 3；Pure accounting, no timer instances *)

(* === 段 1 · 输入校验与量程闸 === *)
uCode := 16#0000;                       // 每拍清码，条件不满足再置（可达清零）/ Clear codes each scan
bDimOk := (fFilmLenM = fFilmLenM) AND (fFilmWidthM = fFilmWidthM) AND (fThickUm = fThickUm)
          AND (fDensityGcc = fDensityGcc)                                          // NaN 自反判据 / NaN reflexivity
          AND (fFilmLenM > fEps) AND (fFilmWidthM > fEps)                          // 长/宽正域闸 / Length and width gate
          AND (fThickUm > fEps) AND (fDensityGcc > fEps)                           // 厚/密正域闸 / Thickness and density gate
          AND (ABS(fDensityGcc) < 1.0E308);                                        // Inf 上限判据 / Inf limit
bCntOk := (nPackCnt >= 1) AND (fPriceYuanKg >= 0.0) AND (fPriceYuanKg = fPriceYuanKg);
                                        // 包数下限闸 + 价格非负闸 / Count and price gates
IF NOT bDimOk OR NOT bCntOk THEN
    uCode := 16#005D;                   // 故障级：域外，核算冻结 / Fault: domain invalid, frozen
END_IF

(* === 段 2 · 主逻辑：量纲链换算 === *)
IF bDimOk THEN
    fDenGcc3 := fDensityGcc * DL_SFC_G2KG;              // 密度 SI 换算 [kg/m³] / Density to SI
    fThickM  := fThickUm * DL_SFC_UM2M;                 // 厚度 SI 换算 [m] / Thickness to SI
    fPerPackKg := fFilmLenM * fFilmWidthM * fThickM * fDenGcc3;     // 单包重量 [kg] / Weight per pack
END_IF

(* === 段 3 · 输出映射与故障码 === *)
    IF bLedgerClr THEN                  (* 台账清零（可达复位路径）/ Ledger clear, reachable reset *)
        fTotalKgAcc := 0.0;             (* 清重量累计 / Clear weight ledger *)
        fCostYuanAcc := 0.0;            (* 清成本累计 / Clear cost ledger *)
    END_IF
    IF bDimOk AND bCntOk THEN
        fTotalKg := fPerPackKg * UDINT_TO_LREAL(INT_TO_UDINT(nPackCnt));    // 产量口径对齐 / Align with pack count
        fCostYuan := fTotalKg * fPriceYuanKg;               // 总成本 [元] / Total cost
        fCostPerPackYn := fCostYuan / UDINT_TO_LREAL(INT_TO_UDINT(nPackCnt));   // 单包成本，包数 ≥1 已闸 / Cost per pack
        fTotalKgAcc := fTotalKgAcc + fTotalKg;      (* 台账累加本拍总耗 / Accumulate the ledger *)
        fCostYuanAcc := fCostYuanAcc + fCostYuan;   (* 台账累加本拍成本 / Accumulate the ledger *)
        IF nCycles < DL_SFC_WRAP THEN
        nCycles := nCycles + 1;         // 有效核算计数，防回卷 / Count valid calculations
    END_IF
ELSIF NOT bDimOk THEN
    fPerPackKg := 0.0;                  // 域外输出安全零 / Safe zero on fault
    fTotalKg := 0.0;
    fCostYuan := 0.0;
    fCostPerPackYn := 0.0;
END_IF
bError := (uCode <> 16#0000);           // 故障标志配对 / Fault flag paired
uErrorId := WORD_TO_UDINT(uCode);       // 码位单点写入（16#0000_005D 形态）/ Single write point
END_FUNCTION_BLOCK

(* ---- FB_DL_SignalStatistics.st ---- *)
(*==============================================================================
 * 组件名称 (Component)  : FB_DL_SignalStatistics
 * 所属子库 (Sublibrary) : DL_MathData
 * 当前版本 (Version)    : 1.0.0
 * 兼容性   (Platform)   : CODESYS 3.5 / TwinCAT 3 / 汇川 InoProShop / Machine Expert
 *                         仅依赖 Standard.library（ABS / MIN / SQRT），无厂商方言
 * 功能描述 (Function)   : 采样流实时统计分析器，滑动窗口（2..64）内输出均值、
 *                         最小值、最大值、峰峰值、样本方差、样本标准差、样本数
 *                         七元组。用于 PID 整定前的噪声评估、SPC 过程能力分析、
 *                         称重稳定性判定、振动烈度监视。
 *                         方差用两遍法：第一遍求均值，第二遍累加离差平方和。
 * 本文件内含       : E_DL_StatState（枚举，归属本组件）
 *                    FB_DL_SignalStatistics（功能块主体）
 * 开源溯源 (Origin)     : 原创实现（参考西门子 LGF 数学组的统计函数分类方式
 *                         与 OSCAT Basic 的标准差/方差/极差行为定义（EPL-2.0）；
 *                         OSCAT 为整数组一次计算，本块为流式窗口，语义不同，
 *                         clean-room 编写，未复制任何源码）。
 * 依赖     (Depends)    : 无 DL_ 内部依赖
 * 红线自检 (Redline)    : R1 ✓ 零全局变量表与外部变量引用 ｜ R2 ✓ 零物理 IO 地址直写
 *                         R3 ✓ 纯 IEC 61131-3，累加用 LREAL 并显式转回 REAL
 *                         R4 ✓ 窗口钳位 + 环形取数正数化取模 + 除零前判 n<2 + NaN 跳过
 *                         R5 ✓ 全变量中英双语同行注释 ｜ R6 ✓ ENUM + CASE + ELSE 兜底
 *                         R7 N/A（无定时器/边沿实例）
 *
 * 【方差公式披露 / Variance-formula disclosure（边界 B1）】
 *   **必须两遍法**。"平方和减均值平方"（E[x²] − E[x]²）在均值远大于标准差时
 *   （如 1000.0 ± 0.01）因灾难性抵消会算出负方差或 0，是 SPC 场景的
 *   经典事故。本块两遍遍历，多一遍 O(n) 换数值安全。
 *
 * 【样本方差口径 / Sample-variance convention（边界 B4）】
 *   用 n−1 分母（样本方差），因为 PLC 拿到的是抽样：与 Excel 的 STDEV.S
 *   一致，不是 STDEV.P。n < 2 时不做除法，方差与标准差输出 0 并置
 *   16#0002_0009（样本不足，瞬时码）。
 *
 * 【极值重算披露 / Extrema-recalc disclosure（边界 B3）】
 *   窗口滑动时若滑出的样本恰为当前极值，增量维护会残留旧极值；
 *   本块每拍随均值遍历一并重算极值（64 点代价可接受），简单且可验证。
 *
 * 【数值类型披露 / Numeric-type disclosure（边界 B7）】
 *   累加与离差用 LREAL（仅为抗累加误差），输出显式转回 REAL，
 *   与现场模拟量量程口径一致。
 *
 * 【验收向量 / Acceptance vectors】
 *   V1  窗口 8，序列 2,4,4,4,5,5,7,9 → fMean = 5.0、fMin = 2、fMax = 9、
 *       fRange = 7、fVariance = 32/7 ≈ 4.5714、fStdDev ≈ 2.1381
 *   V2  单样本 42 → fMean = 42、fVariance = 0、bStatValid = FALSE、16#0002_0009
 *   V3  8 个 3.0 → fMean = 3.0、fVariance = 0.0（非负、非 NaN，边界 B5）
 *   V4  1000.0 与 1000.01 交替 8 个 → 方差 ≈ 2.857e-5（远大于 0，
 *       证明两遍法未发生灾难性抵消）
 *   V5  窗口设 65 → 生效 64、16#0001_0001
 *   V6  V1 后 bClear 一拍 → nCount = 0、bValid = FALSE
 * 修订历史 (Revision)   :
 *   2026-11-14  v1.0.0  首版入库（Phase 1 收口批次 · R3）
 *============================================================================*)
TYPE E_DL_StatState :
(
    eEmpty   := 0,    // 无样本 / No samples yet
    eFilling := 10,   // 样本不足窗口，均值与极值已可用 / Filling, mean and extrema already valid
    eReady   := 20,   // 窗口已满，全部统计量有效 / Window full, all statistics valid
    eFault   := 99    // 参数事件当拍（已钳位，下拍恢复）/ Parameter event scan, clamped, recovers next scan
);
END_TYPE

FUNCTION_BLOCK FB_DL_SignalStatistics
VAR_INPUT
    fIn       : REAL;                      // 采样输入 [EU] / Sample input [EU]
    bSample   : BOOL := TRUE;              // TRUE = 本拍采一个样本（给单周期脉冲即按需采样） / TRUE: take one sample this scan
    nWindow   : INT   := 32;               // 窗口长度，2..64，越界自动钳位 / Window length, range 2..64, clamped
    bClear    : BOOL;                      // TRUE：清空窗口重新统计 / TRUE: clear window and restart
END_VAR
VAR_OUTPUT
    fMean     : REAL;                      // 窗口均值 [EU] / Window mean [EU]
    fMin      : REAL;                      // 窗口最小值 [EU] / Window minimum [EU]
    fMax      : REAL;                      // 窗口最大值 [EU] / Window maximum [EU]
    fRange    : REAL;                      // 峰峰值 fMax − fMin [EU] / Peak-to-peak [EU]
    fVariance : REAL;                      // 样本方差（n−1）[EU²] / Sample variance [EU^2]
    fStdDev   : REAL;                      // 样本标准差 [EU] / Sample standard deviation [EU]
    nCount    : INT;                       // 当前有效样本数 [个] / Valid sample count
    bValid    : BOOL;                      // 至少有 1 个样本（均值/极值有效） / At least one sample, mean valid
    bStatValid: BOOL;                      // 方差/标准差有效（n ≥ 2） / Variance valid, needs n ≥ 2
    uErrorId  : UDINT;                     // 故障码，0 = 无故障（本块码均为瞬时，逐拍重算） / Error code, transient, recomputed every scan
    eState    : E_DL_StatState;            // 当前状态（供诊断） / Current state for diagnostics
END_VAR
VAR
    afWindow  : ARRAY[0..63] OF REAL;      // 环形样本窗 [EU] / Circular sample window [EU]
    nWrite    : INT;                       // 写指针，值域 0..63 / Write index, range 0..63
    nCountInt : INT;                       // 有效样本数（内部） / Internal valid sample count
    nWinEff   : INT;                       // 生效窗口（钳位后） / Effective window after clamping
    nLastWin  : INT;                       // 上拍生效窗口（变更检测，触发整窗重填） / Previous window, change forces refill
    nK        : INT;                       // 遍历索引 / Traversal index
    nIdx      : INT;                       // 环形取数换算下标 / Resolved ring index
    fSum      : LREAL;                     // 均值累加器（宽类型抗漂移） / Sum accumulator for the mean
    fMeanInt  : LREAL;                     // 均值中间量 / Mean intermediate
    fVarAcc   : LREAL;                     // 离差平方和 / Sum of squared deviations
    fTmp      : LREAL;                     // 单点离差 / Single deviation
    fMinInt   : REAL;                      // 本拍重算的窗口最小值 [EU] / Recomputed window minimum [EU]
    fMaxInt   : REAL;                      // 本拍重算的窗口最大值 [EU] / Recomputed window maximum [EU]
    nGuard    : INT;                       // 遍历防死锁计数器 / Traversal guard counter
    bParamEvt : BOOL;                      // 本拍发生参数钳位或窗口变更 / Parameter clamp or window change this scan
    eStateInt : E_DL_StatState;            // 内部状态机当前态 / Internal state machine state
END_VAR
VAR CONSTANT
    DL_STAT_WIN_MIN : INT   := 2;         // 最小窗口（方差需 n ≥ 2） / Minimum window, variance needs n ≥ 2
    DL_STAT_WIN_MAX : INT   := 64;        // 最大窗口（= 数组维度） / Maximum window, equals the array dimension
    DL_STAT_CAP     : INT   := 64;        // 环形容量，必须与数组维度严格一致 / Ring capacity, must match the array
    DL_STAT_GUARD   : INT   := 256;       // 单遍遍历防死锁上限（容量 × 4） / Traversal guard limit, capacity times 4
    DL_STAT_INF_LIM : REAL  := 1.0E30;    // 非有限值判据阈值（超此视为 Inf） / Infinity threshold for non-finite detection
END_VAR

(*------------------------------------------------------------------------------
 * 段 1｜故障码本周期清零：本块故障码全部为瞬时码，逐拍重算
 *      Error code cleared every scan: all codes are transient
 *-----------------------------------------------------------------------------*)
uErrorId  := 16#0000_0000;
bParamEvt := FALSE;

(*------------------------------------------------------------------------------
 * 段 2｜窗口规整：越界钳位，只在本拍置码不刷屏
 *      Window normalization: clamp, code set only on the event scan
 *-----------------------------------------------------------------------------*)
nWinEff := nWindow;
IF nWinEff < DL_STAT_WIN_MIN THEN
    nWinEff  := DL_STAT_WIN_MIN;
    bParamEvt := TRUE;
END_IF
IF nWinEff > DL_STAT_WIN_MAX THEN
    nWinEff  := DL_STAT_WIN_MAX;
    bParamEvt := TRUE;
END_IF
IF bParamEvt THEN
    uErrorId := 16#0001_0001;           // 窗口非法已钳位 / Window invalid, clamped
END_IF

(*------------------------------------------------------------------------------
 * 段 3｜窗口变更检测（R14 语义参数变更）：生效窗口与上拍不同 → 整窗作废
 *      Window change detection: effective window differs, whole window voided
 *-----------------------------------------------------------------------------*)
IF nWinEff <> nLastWin THEN
    nCountInt := 0;
    nWrite    := 0;
    IF nLastWin <> 0 THEN               // 上电首扫不算参数事件 / Power-up first scan is not a parameter event
        uErrorId  := 16#0001_0001;      // 窗口变更触发重填 / Window change forces refill
        bParamEvt := TRUE;
    END_IF
END_IF
nLastWin := nWinEff;

(*------------------------------------------------------------------------------
 * 段 4｜清空：电平触发，先于采样处理
 *      Clear: level-triggered, handled before sampling
 *-----------------------------------------------------------------------------*)
IF bClear THEN
    nCountInt := 0;
    nWrite    := 0;
END_IF

(*------------------------------------------------------------------------------
 * 段 5｜采样（边界：NaN/Inf 跳过不入窗）
 *      Sampling: NaN or Inf samples are skipped, never stored
 *-----------------------------------------------------------------------------*)
IF bSample THEN
    IF (fIn <> fIn) OR (ABS(fIn) > DL_STAT_INF_LIM) THEN
        uErrorId := 16#0001_0006;       // 样本非有限值已跳过 / Non-finite sample skipped
    ELSIF (nWrite >= 0) AND (nWrite < DL_STAT_CAP) THEN
        (* 写指针双检（红线 R4）：MOD 已保证范围，仍显式兜底防越界写 *)
        (* Write index double check: explicit guard besides MOD *)
        afWindow[nWrite] := fIn;
        nWrite    := (nWrite + 1) MOD DL_STAT_CAP;
        nCountInt := MIN(nCountInt + 1, nWinEff);
    END_IF
END_IF

(*------------------------------------------------------------------------------
 * 段 6｜第一遍：均值与极值（边界 B3 极值每拍重算，边界 B7 宽类型累加）
 *      Pass 1: mean and extrema, extrema recomputed every scan
 *-----------------------------------------------------------------------------*)
IF nCountInt > 0 THEN

    fSum   := 0.0;
    nGuard := 0;
    FOR nK := 0 TO (nCountInt - 1) DO
        nGuard := nGuard + 1;
        IF nGuard > DL_STAT_GUARD THEN
            uErrorId := 16#0001_0004;   // 遍历保护触发，保留已算部分 / Traversal guard tripped, partial result kept
            EXIT;
        END_IF
        (* 正数化取模：先加两倍容量再取模，规避负数取模的平台差异 *)
        (* Positive modulo: add twice the capacity before MOD, platform-safe *)
        nIdx := (nWrite - 1 - nK + DL_STAT_CAP * 2) MOD DL_STAT_CAP;
        IF (nIdx < 0) OR (nIdx >= DL_STAT_CAP) THEN
            uErrorId := 16#0001_0004;   // 下标越界兜底（红线 R4） / Index guard fallback
            EXIT;
        END_IF
        fSum := fSum + afWindow[nIdx];
        IF nK = 0 THEN
            fMinInt := afWindow[nIdx];  // 首样本作极值哨兵 / First sample seeds both extrema
            fMaxInt := afWindow[nIdx];
        ELSE
            IF afWindow[nIdx] < fMinInt THEN
                fMinInt := afWindow[nIdx];
            END_IF
            IF afWindow[nIdx] > fMaxInt THEN
                fMaxInt := afWindow[nIdx];
            END_IF
        END_IF
    END_FOR;

    fMeanInt := fSum / INT_TO_LREAL(nCountInt);  // nCountInt > 0 已由段 6 入口保证 / Guaranteed positive at this point

    (*------------------------------------------------------------------------------
     * 段 7｜第二遍：离差平方和（边界 B1 两遍法，边界 B2 除零前判 n < 2）
     *      Pass 2: squared deviations, division guarded by n < 2
     *-----------------------------------------------------------------------------*)
    IF nCountInt >= 2 THEN

        fVarAcc := 0.0;
        nGuard  := 0;
        FOR nK := 0 TO (nCountInt - 1) DO
            nGuard := nGuard + 1;
            IF nGuard > DL_STAT_GUARD THEN
                uErrorId := 16#0001_0004;   // 遍历保护触发 / Traversal guard tripped
                EXIT;
            END_IF
            nIdx := (nWrite - 1 - nK + DL_STAT_CAP * 2) MOD DL_STAT_CAP;
            IF (nIdx < 0) OR (nIdx >= DL_STAT_CAP) THEN
                uErrorId := 16#0001_0004;   // 下标越界兜底（红线 R4） / Index guard fallback
                EXIT;
            END_IF
            fTmp    := afWindow[nIdx] - fMeanInt;
            fVarAcc := fVarAcc + fTmp * fTmp;
        END_FOR;

        fVarAcc := fVarAcc / INT_TO_LREAL(nCountInt - 1);  // n ≥ 2 已判，分母 ≥ 1 / Guarded, denominator ≥ 1

        (* 负方差钳位：浮点舍入可能给出 -1e-20 量级的负零，必须归零 *)
        (* Negative variance clamp: rounding may yield tiny negative zeros *)
        IF fVarAcc < 0.0 THEN
            fVarAcc := 0.0;
        END_IF

    ELSE
        fVarAcc   := 0.0;
        uErrorId  := 16#0002_0009;      // 样本不足（N < 2，方差无定义）/ Too few samples for variance
    END_IF

ELSE
    fSum      := 0.0;
    fMeanInt  := 0.0;
    fVarAcc   := 0.0;
    fMinInt   := 0.0;
    fMaxInt   := 0.0;
END_IF

(*------------------------------------------------------------------------------
 * 段 8｜派生统计量：标准差与峰峰值，显式 LREAL_TO_REAL 回写
 *      Derived statistics: standard deviation and peak-to-peak, explicit casts
 *-----------------------------------------------------------------------------*)
fMean     := LREAL_TO_REAL(fMeanInt);
fVariance := LREAL_TO_REAL(fVarAcc);
fStdDev   := LREAL_TO_REAL(SQRT(fVarAcc));
fMin      := fMinInt;
fMax      := fMaxInt;
fRange    := fMaxInt - fMinInt;

(*------------------------------------------------------------------------------
 * 段 9｜状态派生与主状态机（红线 R6）：ENUM + CASE + ELSE 兜底
 *      State derivation and main state machine with ELSE fallback
 *-----------------------------------------------------------------------------*)
IF bParamEvt THEN
    eStateInt := E_DL_StatState.eFault;
ELSIF nCountInt <= 0 THEN
    eStateInt := E_DL_StatState.eEmpty;
ELSIF nCountInt < nWinEff THEN
    eStateInt := E_DL_StatState.eFilling;
ELSE
    eStateInt := E_DL_StatState.eReady;
END_IF

CASE eStateInt OF

    E_DL_StatState.eEmpty:
        (* 无样本：统计量保持段 8 的零值，bValid 由段 10 置 FALSE / No samples *)

    E_DL_StatState.eFilling:
        (* 填充中：均值/极值已有效，方差是否有效由 bStatValid 表达（边界 B4） *)
        (* Filling: mean valid, variance validity carried by bStatValid *)

    E_DL_StatState.eReady:
        (* 就绪：全部统计量有效 / Ready: all statistics valid *)

    E_DL_StatState.eFault:
        (* 参数事件当拍：参数已修正、下拍恢复，不锁存 / Event scan, recovers next scan *)

    ELSE
        (* 非法状态一律回故障态并置码（红线 R6） *)
        (* Illegal state falls back to fault with a code *)
        eStateInt := E_DL_StatState.eFault;
        uErrorId  := 16#0001_0005;

END_CASE

(*------------------------------------------------------------------------------
 * 段 10｜输出单一出口：有效标志由计数派生
 *      Single output exit: validity flags derived from the count
 *-----------------------------------------------------------------------------*)
nCount     := nCountInt;
bValid     := (nCountInt > 0);
bStatValid := (nCountInt >= 2);
eState     := eStateInt;
END_FUNCTION_BLOCK

(* ---- FB_DL_SkewKurtosisCalc.st ---- *)
(*
  ==================================================================
  组件名 Component  : FB_DL_SkewKurtosisCalc
  分类   Category   : DL_MathData
  复杂度 Complexity  : cx5
  版本   Version    : 1.0.0
  功能   Purpose    : 在线偏度 / 峰度统计。Welford 高阶矩递推（单遍、数值稳
                      定），输出均值 / 偏度 g1 / 超额峰度 g2；非有限样本剔除
                      并计数；样本数不足或方差退化时统计量出口归零并降
                      bValid。与 StdDevOnline / CovarOnline 同族补口（高阶矩）。
  来源   Source     : t2-1-lgf-math（统计族待挖项）
  溯源   Origin     : Welford 递推为公开数值算法（教学资料），clean-room 自研
                      实现；未复制任何厂商私有库源码。
  平台   Platform   : 纯 IEC 61131-3（Standard.library: R_TRIG / SQRT，无私有库）
  分工声明 Split     : 与 FB_DL_StdDevOnline / FB_DL_CovarOnline 分工——StdDev
                      为一阶 / 二阶矩在线统计，Covar 为双序列协方差；本件补
                      三阶 / 四阶矩（偏度与峰度），不做双序列与回归。
  作者   Author     : 道莅代码库 · PLC 编程专家（R58）
  ------------------------------------------------------------------
  边界 Boundary     :
                      一 有效样本数 nCnt ≥ 4 才出偏度 / 峰度（四阶矩稳定性
                      门槛，不足时出口归零 + bValid = FALSE，信息级降级）；
                      二 二阶矩 _lrM2 ≤ 1E-300 视为方差退化：偏度 / 峰度归零
                      （等值序列无形状信息），bValid 仍为 TRUE；
                      三 非有限样本（NaN 自反 / Inf 差值自减双判据）剔除计
                      数 nNanCnt，不参与递推；
                      四 复位沿作用域：清累计量 / 清出口（两项逐项声明），
                      首扫执行与复位沿同款初始化（R310 _bInit）；
                      五 无全局变量、无外部变量声明、无物理地址寻址。
  修订记录 Revision  :
    2026-11-21  v1.0.0  R58 首版（批 1 · 序号 4）
  ==================================================================
*)

FUNCTION_BLOCK FB_DL_SkewKurtosisCalc
VAR_INPUT
    fX     : LREAL := 0.0;  // 样本输入 [工程单位] / the sample input [engineering unit]
    bSample: BOOL := FALSE; // 样本有效电平，TRUE = 本拍样本参与统计 [-] / the sample valid level, true includes this scan
    bReset : BOOL := FALSE; // 复位上升沿清全部统计 [-] / reset rising edge clears all statistics
END_VAR
VAR_OUTPUT
    fMean   : LREAL := 0.0; // 均值出口 [工程单位] / the mean outlet [engineering unit]
    fSkew   : LREAL := 0.0; // 偏度出口 g1（无量纲）/ the skewness outlet, dimensionless
    fKurt   : LREAL := 0.0; // 超额峰度出口 g2（无量纲，正态为 0）/ the excess kurtosis outlet, dimensionless, zero for normal
    nCnt    : UDINT := 0;   // 有效样本数 [个] / the valid sample count
    nNanCnt : UDINT := 0;   // 剔除的非有限样本数 [个] / the excluded non finite sample count
    bValid  : BOOL := FALSE; // 统计量有效（nCnt ≥ 4 且形状可算）[-] / the statistics valid flag
END_VAR
VAR
    rtReset : R_TRIG; // 复位沿检测，段 0 无条件刷新 / the reset edge, refreshed unconditionally
    _bInit  : BOOL := FALSE; // 首扫初始化完成标志（R310）/ the first scan flag
    _lrM2   : LREAL := 0.0;  // 二阶中心矩累加器（Welford M2）[工程单位平方] / the second central moment accumulator [unit squared]
    _lrM3   : LREAL := 0.0;  // 三阶中心矩累加器（Welford M3）[工程单位立方] / the third central moment accumulator [unit cubed]
    _lrM4   : LREAL := 0.0;  // 四阶中心矩累加器（Welford M4）[工程单位四次方] / the fourth central moment accumulator [unit to the fourth]
    _lrN    : LREAL;         // 当前样本数实数副本 [个] / the current count as a real [count]
    _lrDlt  : LREAL;         // 本拍偏差 [工程单位] / the delta this scan [engineering unit]
    _lrDltN : LREAL;         // 归一偏差 [工程单位] / the normalized delta [engineering unit]
    _lrD2   : LREAL;         // 归一偏差平方 [工程单位平方] / the normalized delta squared
    _lrT1   : LREAL;         // Welford 一阶项 [工程单位平方] / the Welford first term
    _lrSd   : LREAL;         // 标准差工作量 [工程单位] / the standard deviation work value
END_VAR
VAR CONSTANT
    DL_SK_MINCNT : UDINT := 4;          // 统计量出口最小样本数 [个]（边界一）/ the minimum sample count for the shape outlets
    DL_SK_TINY   : LREAL := 1.0E-300;   // 方差退化阈值 [工程单位平方]（边界二）/ the variance degeneration threshold
    DL_SK_CNTMAX : UDINT := 4294967294; // 样本数累加钳定界 [个]，防 UDINT 回绕 / the count clamp against a wrap
END_VAR

// 段 0｜沿检测无条件周期刷新（禁入分支）/ segment 0, the unconditional refresh
rtReset(CLK := bReset); // 复位沿 / the reset edge

// 段 1｜首扫初始化（R310）：与复位沿同款初始化块 / segment 1, the first scan init, the same block as the reset edge
IF NOT _bInit THEN // 首扫一拍 / the first scan
    _bInit := TRUE; // 置首扫标志 / raise the first scan flag
    _lrM2 := 0.0; // 二阶矩清零 / clear M2
    _lrM3 := 0.0; // 三阶矩清零 / clear M3
    _lrM4 := 0.0; // 四阶矩清零 / clear M4
END_IF

// 段 2｜复位沿作用域：清累计量 / 清出口（两项逐项声明，边界四）/ segment 2, the reset edge scope
IF rtReset.Q THEN // 复位沿 / the reset edge
    nCnt := 0; // 作用域一：清有效样本数 / scope one, clear the count
    nNanCnt := 0; // 作用域一：清剔除计数 / scope one, clear the excluded count
    fMean := 0.0; // 作用域一：清均值出口 / scope one, clear the mean
    _lrM2 := 0.0; // 作用域一：清二阶矩 / scope one, clear M2
    _lrM3 := 0.0; // 作用域一：清三阶矩 / scope one, clear M3
    _lrM4 := 0.0; // 作用域一：清四阶矩 / scope one, clear M4
    fSkew := 0.0; // 作用域二：清偏度出口 / scope two, clear the skewness
    fKurt := 0.0; // 作用域二：清峰度出口 / scope two, clear the kurtosis
    bValid := FALSE; // 作用域二：清有效标志 / scope two, clear the valid flag
END_IF

// 段 3｜样本受理与非有限剔除（边界三）/ segment 3, the sample admission and the non finite exclusion
IF bSample THEN // 本拍有样本 / a sample this scan
    IF (fX = fX) AND ((fX - fX) = (fX - fX)) THEN // 有限样本双判据通过（R79）/ a finite sample by the dual verdicts
        IF nCnt < DL_SK_CNTMAX THEN // 计数未到钳定界 / below the count clamp
            _lrN := UDINT_TO_LREAL(nCnt) + 1.0; // 新样本数实数副本（≥1，除子安全）/ the new count as a real
            _lrDlt := fX - fMean; // 本拍偏差 / the delta
            _lrDltN := _lrDlt / _lrN; // 归一偏差（除子已证 ≥1）/ the normalized delta
            _lrD2 := _lrDltN * _lrDltN; // 归一偏差平方 / the normalized delta squared
            _lrT1 := _lrDlt * _lrDltN * (_lrN - 1.0); // Welford 一阶项 / the Welford first term
            _lrM4 := _lrM4 + _lrT1 * _lrD2 * (_lrN * _lrN - 3.0 * _lrN + 3.0) + 6.0 * _lrD2 * _lrM2 - 4.0 * _lrDltN * _lrM3; // 四阶矩递推 / the fourth moment recursion
            _lrM3 := _lrM3 + _lrT1 * _lrDltN * (_lrN - 2.0) - 3.0 * _lrDltN * _lrM2; // 三阶矩递推 / the third moment recursion
            _lrM2 := _lrM2 + _lrT1; // 二阶矩递推 / the second moment recursion
            fMean := fMean + _lrDltN; // 均值推进 / advance the mean
            nCnt := nCnt + 1; // 有效样本数推进 / advance the count
        ELSE // 已在钳定界（防回绕，拒绝新样本计数推进）/ at the clamp, the count frozen
            nCnt := DL_SK_CNTMAX; // 钳定保持 / hold at the clamp
        END_IF
    ELSE // 非有限样本剔除（边界三）/ a non finite sample excluded
        IF nNanCnt < DL_SK_CNTMAX THEN // 剔除计数防回绕 / the exclusion count wrap guard
            nNanCnt := nNanCnt + 1; // 剔除计数推进 / advance the excluded count
        END_IF
    END_IF
END_IF

// 段 4｜形状统计量出口计算（样本数与方差双门槛，边界一二）/ segment 4, the shape outlets
bValid := (nCnt >= DL_SK_MINCNT); // 有效标志：样本数门槛 / the valid flag, the count gate
IF bValid AND (_lrM2 > DL_SK_TINY) THEN // 样本足且方差未退化 / enough samples and a live variance
    _lrSd := SQRT(_lrM2 / UDINT_TO_LREAL(nCnt)); // 标准差工作量（除子已证 ≥4）/ the standard deviation work value
    fSkew := SQRT(UDINT_TO_LREAL(nCnt)) * _lrM3 / (_lrM2 * SQRT(_lrM2)); // g1 = √n·M3 / M2^1.5（除子已证 >0）/ the skewness, the divisor proven positive
    fKurt := UDINT_TO_LREAL(nCnt) * _lrM4 / (_lrM2 * _lrM2) - 3.0; // g2 = n·M4 / M2² - 3（除子已证 >0）/ the excess kurtosis, the divisor proven positive
ELSE // 不足或退化：出口归零（信息级降级，不置故障）/ short or degenerate, the outlets zeroed
    fSkew := 0.0; // 偏度归零 / zero the skewness
    fKurt := 0.0; // 峰度归零 / zero the kurtosis
END_IF

// 段 5｜出口非有限复检兜底（防御纵深，正常路径不可达）/ segment 5, the outlet recheck as defense in depth
IF (fSkew <> fSkew) OR ((fSkew - fSkew) <> (fSkew - fSkew)) THEN // 偏度非有限 / a non finite skewness
    fSkew := 0.0; // 归零兜底 / zero the outlet
    bValid := FALSE; // 降有效标志 / drop the valid flag
END_IF
IF (fKurt <> fKurt) OR ((fKurt - fKurt) <> (fKurt - fKurt)) THEN // 峰度非有限 / a non finite kurtosis
    fKurt := 0.0; // 归零兜底 / zero the outlet
    bValid := FALSE; // 降有效标志 / drop the valid flag
END_IF
END_FUNCTION_BLOCK

(* ---- FB_DL_SlurryViscosityComp.st ---- *)
(*
  Component : FB_DL_SlurryViscosityComp
  Category  : DL_MathData
  Type      : FB
  Version   : 1.0.2
  CodeSeg   : 16#02_3_5C
  Summary   : 浆料粘度温度补偿换算：温-粘标定曲线查表线性插值，输出归一到参考温度的补偿后粘度。
              Slurry viscosity temperature compensation: lookup curve linear interpolation, output normalized to reference temperature.
  溯源声明  : 道莅自研 clean-room
  边界安全  : 温度物理域闸（> -273.15 degC，非有限 NaN/Inf 拦截）；粘度正域闸（> 0，防负值换算）；
              曲线点数域闸（2..8，防数组越界访问）；插值端点钳制（域外温度取边界因子并置 xClamped）；
              插值分母（节点温差）先判容差再除，防除零；全浮点比较带 fEps 容差。
  复用      : 无
  修订历史  : v1.0.2（R34 返修）改动点：① bRun=FALSE 分支改为「冻结保持末次有效粘度 + 置 bDegraded := TRUE」，
              禁输出 0 或未定义值；② xClamped 与钳制判据同源赋值（每拍先清零，仅端点钳制时置 TRUE），
              名实相符且不再在无效态残留旧值。接口仅新增 bDegraded 一个输出引脚，其余引脚与顺序一字不动。
              v1.0.0 首版入库。
  降级语义  : bDegraded = TRUE 表示输出为末次有效值的冻结副本（非本拍换算结果），HMI 需标注数据陈旧。
*)

FUNCTION_BLOCK FB_DL_SlurryViscosityComp
VAR_INPUT
    bRun          : BOOL;              (* 换算使能，假则输出冻结 · Enable, FALSE freezes outputs *)
    fTempC        : LREAL;             (* 浆料实测温度 [degC] · Measured slurry temperature *)
    fViscMeasMpas : LREAL;             (* 实测粘度 [mPa·s] · Measured viscosity *)
    fTRefC        : LREAL := 25.0;     (* 参考温度 [degC]，补偿归一基准 · Reference temperature *)
    aCurveTc      : ARRAY[1..8] OF LREAL := [5.0, 15.0, 25.0, 35.0, 45.0, 55.0, 65.0, 75.0];
                                       (* 曲线温度节点 [degC]，升序标定 · Curve temperature nodes, ascending *)
    aCurveK       : ARRAY[1..8] OF LREAL := [1.60, 1.30, 1.00, 0.80, 0.65, 0.54, 0.46, 0.40];
                                       (* 各节点补偿因子 [比值] · Compensation factor per node *)
    nPts          : INT := 8;          (* 有效点数 [点]，域 2 到 8 · Valid point count *)
    fEps          : LREAL := 1.0E-6;   (* 浮点判零容差 [实数域] · Floating zero tolerance *)
END_VAR
VAR_OUTPUT
    fViscCompMpas : LREAL;             (* 补偿后粘度 [mPa·s]，归一到参考温度 · Compensated viscosity at reference *)
    fFactorNow    : LREAL;             (* 当前温度补偿因子 [比值] · Factor at current temperature *)
    fFactorRef    : LREAL;             (* 参考温度补偿因子 [比值] · Factor at reference temperature *)
    xClamped      : BOOL;              (* 端点钳制标志 [开关] · Endpoint clamp flag *)
    bError        : BOOL;              (* 故障标志，与故障码配对 · Fault flag paired with codes *)
    uErrorId      : UDINT;             (* 事件码 16#0000_005C，0 无事件 · Event code *)
    bDegraded     : BOOL;              (* v1.0.2 新增：降级标志，TRUE = 输出为末次有效值冻结副本 · Degraded flag, TRUE = frozen last-good output *)
END_VAR
VAR
    uCode   : WORD;    (* 码位暂存，每拍重算 [码] · Code staging, recomputed per scan *)
    bSigOk  : BOOL;    (* 输入有效标志 · Input validity flag *)
    bTblOk  : BOOL;    (* 曲线点数域标志 · Table point-count validity *)
    bRefOk  : BOOL;    (* 参考温度插值有效标志 · Reference interpolation validity *)
    nSeg    : INT;     (* 命中段下标 [索引] · Hit segment index *)
    nI      : INT;     (* 查表循环下标 [索引] · Table loop index *)
    fDen    : LREAL;   (* 插值分母（节点温差）[degC] · Interpolation denominator *)
    nCycles : UDINT;   (* 有效换算拍计数 [拍]，防回卷 · Valid conversion count with wrap guard *)
END_VAR
VAR CONSTANT
    DL_SVC_ABS0 : LREAL := 273.15;     (* 绝对零度 [degC] · Absolute zero in celsius *)
    DL_SVC_WRAP : UDINT := 4294967290; (* 计数防回卷余量 [拍] · Counter wrap guard *)
END_VAR

(* === 段 0 · 实例刷新 === *)
(* 纯换算件：无 TON/R_TRIG 实例，计数状态见段 3；Pure conversion, no timer instances *)

(* === 段 1 · 输入校验与量程闸 === *)
uCode := 16#0000;                       // 每拍清码，条件不满足再置（可达清零）/ Clear codes each scan
bSigOk := (fTempC = fTempC) AND (fViscMeasMpas = fViscMeasMpas) AND (fTRefC = fTRefC)
          AND (ABS(fTempC) < 1.0E308) AND (ABS(fViscMeasMpas) < 1.0E308)     // NaN 自反 + Inf 上限
          AND (fTempC > (-DL_SVC_ABS0 + fEps))                               // 温度物理域闸 / Physical domain
          AND (fViscMeasMpas > fEps)                                         // 粘度正域闸 / Positive viscosity
          AND (fTRefC > (-DL_SVC_ABS0 + fEps));                              // 参考温度域闸 / Reference domain
bTblOk := (nPts >= 2) AND (nPts <= 8);  // 点数域闸，防数组越界 / Point-count gate
IF NOT bSigOk OR NOT bTblOk THEN
    uCode := 16#005C;                   // 故障级：域外或表无效，换算冻结 / Fault: domain or table invalid
END_IF

(* === 段 2 · 主逻辑：查表线性插值（禁止 IF-ELSE 阶梯硬编码）=== *)
xClamped := FALSE;                      // v1.0.2：每拍先清钳制标志，与钳制判据同源（防无效态残留旧 TRUE）
IF bSigOk AND bTblOk THEN
    IF fTempC <= aCurveTc[1] THEN
        fFactorNow := aCurveK[1];       // 低温端点钳制 / Clamp at the low end
        xClamped := TRUE;
    ELSIF fTempC >= aCurveTc[nPts] THEN
        fFactorNow := aCurveK[nPts];    // 高温端点钳制 / Clamp at the high end
        xClamped := TRUE;
    ELSE
        nSeg := nPts - 1;               // 段下标兜底最后一段 / Default to the last segment
        FOR nI := 1 TO (nPts - 1) DO
            IF fTempC <= aCurveTc[nI + 1] THEN
                nSeg := nI;             // 命中段锁定 / Lock the hit segment
                EXIT;
            END_IF
        END_FOR
        fDen := aCurveTc[nSeg + 1] - aCurveTc[nSeg];    // 分母导出 / Denominator
        IF fDen > fEps THEN             // 防除零闸 / Divide-by-zero gate
            fFactorNow := aCurveK[nSeg] + (aCurveK[nSeg + 1] - aCurveK[nSeg])
                          * (fTempC - aCurveTc[nSeg]) / fDen;   // 线性插值 / Linear interpolation
        ELSE
            fFactorNow := aCurveK[nSeg];    // 退化取左节点因子 / Degenerate to left node
        END_IF
    END_IF
    (* 参考温度因子：同一段插值，参考温度域闸已在段 1 保证 / Same interpolation at the reference *)
    IF fTRefC <= aCurveTc[1] THEN
        fFactorRef := aCurveK[1];       // 参考端点钳制 / Reference clamp low
        bRefOk := TRUE;
    ELSIF fTRefC >= aCurveTc[nPts] THEN
        fFactorRef := aCurveK[nPts];    // 参考端点钳制 / Reference clamp high
        bRefOk := TRUE;
    ELSE
        nSeg := nPts - 1;
        FOR nI := 1 TO (nPts - 1) DO
            IF fTRefC <= aCurveTc[nI + 1] THEN
                nSeg := nI;
                EXIT;
            END_IF
        END_FOR
        fDen := aCurveTc[nSeg + 1] - aCurveTc[nSeg];
        IF fDen > fEps THEN
            fFactorRef := aCurveK[nSeg] + (aCurveK[nSeg + 1] - aCurveK[nSeg])
                          * (fTRefC - aCurveTc[nSeg]) / fDen;
        ELSE
            fFactorRef := aCurveK[nSeg];
        END_IF
        bRefOk := TRUE;                 // 参考插值完成 / Reference interpolation done
    END_IF
END_IF

(* === 段 3 · 输出映射与故障码 === *)
bDegraded := FALSE;                     // v1.0.2：降级标志每拍重算，条件满足再置
IF bRun THEN
    IF bSigOk AND bTblOk THEN
        IF fFactorRef > fEps THEN           // 归一分母防除零 / Normalize denominator gate
            fViscCompMpas := fViscMeasMpas * fFactorNow / fFactorRef;   // 归一补偿粘度 / Compensated viscosity
        END_IF
        IF nCycles < DL_SVC_WRAP THEN
            nCycles := nCycles + 1;         // 有效换算计数，防回卷 / Count valid conversions
        END_IF
    ELSE
        bDegraded := TRUE;                  // 输入域外：输出冻结为末次有效值并标降级
        xClamped := FALSE;                  // 无效态不主张钳制（与钳制判据同源）
    END_IF
ELSE
    bDegraded := TRUE;                      // v1.0.2：bRun=FALSE 冻结保持末次有效粘度，禁输出 0
    xClamped := FALSE;                      // v1.0.2：停算态钳制标志清零，名实相符
END_IF
bError := (uCode <> 16#0000);           // 故障标志配对 / Fault flag paired
uErrorId := WORD_TO_UDINT(uCode);       // 码位单点写入（16#0000_005C 形态）/ Single write point
END_FUNCTION_BLOCK

(* ---- FB_DL_StatsRollingVar.st ---- *)
(*
  ============================================================
  组件名 : FB_DL_StatsRollingVar
  分类   : DL_MathData
  功能   : 定长环形缓冲的滚动方差与滚动标准差，最旧样本先移出再插入新样本
  开源溯源 : internal-design（本轮无外部代码逐行引用）
             参考语义 : 无外部参考
  复杂度 : C2
  版本   : 1.0.0
  ============================================================
  口径说明 : 方差为样本方差（分母 n-1），n 小于二时判无效；浮点误差使方差为负时钳到零。
             环形缓冲容量六十四，满后最旧样本先移出。
             复位沿作用域：清缓冲、清和与平方和、清游标与已填数；不清输出语义定义。
             bEnable 为假时冻结保持——不插入新样本，输出继续按既有缓冲计算。
*)

FUNCTION_BLOCK FB_DL_StatsRollingVar
VAR_INPUT
    rInput  : REAL; // 采样输入值 [工程单位] sample input value [engineering unit]
    bEnable : BOOL; // 采样使能，假为冻结保持 sampling enable, false freezes the buffer
    bReset  : BOOL; // 复位命令，上升沿清空缓冲 reset command clearing the buffer on its rising edge
END_VAR
VAR_OUTPUT
    rVariance : REAL; // 样本方差 [工程单位平方] sample variance [engineering unit squared]
    rStd      : REAL; // 样本标准差 [工程单位] sample standard deviation [engineering unit]
    rMean     : REAL; // 样本均值 [工程单位] sample mean [engineering unit]
    nCount    : INT; // 当前缓冲样本数 [个] buffered sample count [count]
    bValid    : BOOL; // 结果有效标志 result validity flag
END_VAR
VAR CONSTANT
    DL_CAP  : INT := 64; // 缓冲容量 [个] buffer capacity [count]
    DL_LAST : INT := 63; // 缓冲末下标 last buffer index
END_VAR
VAR
    _afBuf  : ARRAY[0..63] OF REAL := [64(0.0)]; // 环形样本缓冲 [工程单位] ring sample buffer [engineering unit]
    _nIdx   : INT := 0; // 写入游标 [个] write cursor [count]
    _nFilled: INT := 0; // 已填样本数 [个] filled sample count [count]
    _rSum   : REAL := 0.0; // 样本和 running sum [engineering unit]
    _rSumSq : REAL := 0.0; // 样本平方和 running sum of squares [engineering unit squared]
    _rVar   : REAL := 0.0; // 方差中间量 [工程单位平方] intermediate variance [engineering unit squared]
    _bInit  : BOOL := FALSE; // 首扫初始化标志 first scan initialisation flag
    i       : INT := 0; // 清缓冲游标 [个] clearing cursor [count]
    rtReset : R_TRIG; // 复位上升沿 reset rising edge
END_VAR

// 段 0｜复位沿实例无条件周期刷新 unconditional cyclic refresh of the reset edge
rtReset(CLK := bReset); // 复位沿刷新 refresh the reset edge
// 段 1｜出口预置 preset the exit
rVariance := 0.0; // 方差预置零 variance preset to zero
rStd := 0.0; // 标准差预置零 deviation preset to zero
rMean := 0.0; // 均值预置零 mean preset to zero
bValid := FALSE; // 计算完成前不认结果 unusable before the calculation
// 段 2｜首扫与复位沿初始化 first scan and reset edge initialisation
IF (NOT _bInit) OR rtReset.Q THEN
    FOR i := 0 TO DL_LAST DO
        _afBuf[i] := 0.0; // 逐槽清零 clear every slot
    END_FOR
    _nIdx := 0; // 游标归零 the cursor returns to zero
    _nFilled := 0; // 已填数归零 the filled count returns to zero
    _rSum := 0.0; // 样本和归零 the running sum returns to zero
    _rSumSq := 0.0; // 平方和归零 the sum of squares returns to zero
    _bInit := TRUE; // 首扫初始化完成 the first scan initialisation is done
END_IF
// 段 3｜采样插入，最旧样本先移出 sample insertion with the oldest leaving first
IF bEnable AND (rInput = rInput) THEN
    _rSum := _rSum - _afBuf[_nIdx]; // 移出最旧值占的和 remove the oldest from the sum
    _rSumSq := _rSumSq - _afBuf[_nIdx] * _afBuf[_nIdx]; // 移出最旧值占的平方和 remove the oldest from the squares
    _afBuf[_nIdx] := rInput; // 新样本写入游标位 write the new sample at the cursor
    _rSum := _rSum + rInput; // 累入新样本 accumulate the new sample
    _rSumSq := _rSumSq + rInput * rInput; // 累入新样本平方 accumulate the new square
    IF _nFilled < DL_CAP THEN
        _nFilled := _nFilled + 1; // 未满时已填数递增 count up while the buffer is not full
    END_IF
    _nIdx := _nIdx + 1; // 游标前进 advance the cursor
    IF _nIdx > DL_LAST THEN
        _nIdx := 0; // 满圈回绕 wrap around
    END_IF
END_IF
// 段 4｜统计量计算 statistics computation
nCount := _nFilled; // 样本数出口 map the buffered count
IF _nFilled >= 2 THEN
    rMean := _rSum / INT_TO_REAL(_nFilled); // 均值，除子为已证正样本数 mean over a proven positive count
    _rVar := (_rSumSq - (_rSum * _rSum) / INT_TO_REAL(_nFilled)) / INT_TO_REAL(_nFilled - 1); // 样本方差 sample variance
    IF _rVar < 0.0 THEN
        _rVar := 0.0; // 浮点误差致负时钳零 clamp a negative value caused by rounding
    END_IF
    rVariance := _rVar; // 方差落定 land the variance
    rStd := SQRT(_rVar); // 标准差为方差开方 the deviation is the square root of the variance
    bValid := TRUE; // 结果可用 result usable
ELSIF _nFilled = 1 THEN
    rMean := _rSum; // 单样本时均值即样本值 a single sample is its own mean
END_IF
END_FUNCTION_BLOCK

(* ---- FB_DL_StatsWelfordVar.st ---- *)
(*==============================================================================
 * 组件名称 : FB_DL_StatsWelfordVar ｜ 子库 : DL_MathData ｜ v1.0.0 ｜ 2026-11-24
 * 平台     : CODESYS 3.5 / TwinCAT 3 / InoProShop / Machine Expert（纯 IEC，无厂商库）
 * 功能简介 : Welford 在线均值/方差累加器 —— 单遍递推，不保存样本、不做减法抵消，
 *            长序列下数值稳定性远优于「先求和再平方和」。递推式：
 *            d = x − mean；mean += d/n；M2 += d·(x − mean)；样本方差 = M2/(n−1)。
 * 契约     : bEnable 按「新样本到达」语义使用 —— 只在上升沿采样一次（内部 R_TRIG），
 *            bEnable 保持为真的多个周期不会重复计入同一值。
 *            bReset 上升沿清零 n / mean / M2（R18 用 R_TRIG，禁电平判据）。
 *            出参 fMean / fVar / fStd / nCount / bValid；n = 1 时 fVar := 0；
 *            bValid 仅在 n ≥ 2（三件套同时可用）为真，均值本身 n = 1 即有效。
 *            非有限样本直接丢弃并置 bRejected（单拍），不污染累加器。
 * 依赖     : 无 DL_ 内部依赖（R16 自足实现）；Standard.library: R_TRIG / ABS / SQRT
 * 错误码   : R297 零码位范式：eErr 恒 0，丢弃以 bRejected 表达
 * 红线自检 : R1 零全局 R2 零%I/%Q R3 纯IEC R4 除零前置（n 自增后才整除）、NaN 自反判据、
 *            无穷上界、负方差兜底 ｜ R5 双语注释 R6 ENUM+CASE+ELSE 兜底
 *            R7 R_TRIG 实例置于 CASE 外无条件周期刷新 ｜ R10 标准转换
 *            R11 全声明行分号 R14 无 PROPERTY R15 标识符零保留字冲突
 *            R18 bReset 走 R_TRIG 上升沿
 * 修订历史 : 2026-11-24 R79-A 首版（统计扩展族 1/8）
 *============================================================================*)
TYPE E_DL_WelfordStage :
(
    eWelfordIdle  := 0,     // 零样本，无均值 / no sample, no mean
    eWelfordAccum := 1,     // 单样本，均值可用方差不可用 / one sample, the mean exists but the variance does not
    eWelfordReady := 2      // 两样本以上，均值方差均可用 / two samples or more, everything is usable
);
END_TYPE

FUNCTION_BLOCK FB_DL_StatsWelfordVar
VAR_INPUT
    bEnable   : BOOL;   // 采样使能，上升沿表示新样本到达 / capture enable, a rising edge marks a new sample
    bReset    : BOOL;   // 复位，上升沿清零全部累加器 / reset, a rising edge clears every accumulator
    fSample   : LREAL;  // 样本值，非有限者被丢弃 [工程单位] / sample value, non finite ones are dropped [engineering unit]
END_VAR
VAR_OUTPUT
    eErr      : UDINT;  // 错误码，零码位范式恒 0 / error id, always zero under the zero-code rule
    bError    : BOOL;   // 故障标志，本件不产生故障级 / fault flag, never raised by this component
    bRejected : BOOL;   // 本拍样本被丢弃（非有限） / TRUE when this cycle sample was dropped
    fMean     : LREAL;  // 在线均值 [工程单位] / running mean [engineering unit]
    fVar      : LREAL;  // 样本方差（n−1 分母），n=1 时为 0 [工程单位²] / sample variance with the n minus one divisor [unit squared]
    fStd      : LREAL;  // 样本标准差 [工程单位] / sample standard deviation [engineering unit]
    nCount    : UDINT;  // 已纳入样本数 [个] / number of accepted samples [count]
    bValid    : BOOL;   // n ≥ 2 时为真，三件套同时可用 / TRUE from two samples on, when all three outputs are usable
    eStage    : E_DL_WelfordStage;  // 累加器阶段 / accumulator stage
END_VAR
VAR CONSTANT
    DL_ONE      : UDINT := 1;           // 无符号一 / unsigned one
    DL_TWO      : UDINT := 2;           // 无符号二，方差可用门槛 / unsigned two, the usable variance threshold
    DL_FIN_LIM  : LREAL := 1.0E308;     // 有限性上界，超过按无穷处置 [工程单位] / finiteness ceiling [engineering unit]
    DL_ZERO_L   : LREAL := 0.0;         // 实数零哨兵 / real zero sentinel
END_VAR
VAR
    rtReset   : R_TRIG; // 复位上升沿检测，无条件周期刷新 / reset rising edge, refreshed every cycle
    rtSample  : R_TRIG; // 采样上升沿检测，无条件周期刷新 / sample rising edge, refreshed every cycle
    nAcc      : UDINT;  // 内部样本计数 / internal sample counter
    fMeanInt  : LREAL;  // 内部均值累加器 [工程单位] / internal mean accumulator [engineering unit]
    fM2       : LREAL;  // 二阶中心矩累加器 M2 [工程单位²] / second central moment accumulator [unit squared]
    fDelta    : LREAL;  // 偏差 d = x − mean [工程单位] / deviation of the new sample [engineering unit]
    fVarInt   : LREAL;  // 方差中间量，负偏时兜底到 0 [工程单位²] / variance interim value, clamped at zero [unit squared]
END_VAR

// 段 1｜沿检测无条件周期刷新（R7）：先刷新，后判定 / segment 1, refresh both edges unconditionally before any test
rtReset(CLK := bReset);
rtSample(CLK := bEnable);

// 段 2｜出口预置：单拍量与码位每拍重算 / segment 2, preset the single cycle outputs
eErr      := 0;             // 零码位范式 / zero-code rule
bError    := FALSE;         // 本件不产生故障级 / this component raises no fault
bRejected := FALSE;         // 本拍未丢弃 / nothing dropped yet

// 段 3｜复位优先：上升沿清 n / mean / M2，不动阶段（阶段在段 5 回落）/ segment 3, reset has priority
IF rtReset.Q THEN
    nAcc     := 0;          // 计数清零 / clear the counter
    fMeanInt := DL_ZERO_L;  // 均值清零 / clear the mean
    fM2      := DL_ZERO_L;  // 二阶矩清零 / clear the second moment
END_IF

// 段 4｜采样：仅上升沿计入，非有限样本丢弃 / segment 4, capture on the rising edge only
IF rtSample.Q THEN
    IF (fSample <> fSample) OR (ABS(fSample) > DL_FIN_LIM) THEN
        bRejected := TRUE;                                  // 非数或无穷，丢弃 / not a number or infinity, dropped
    ELSE
        nAcc     := nAcc + DL_ONE;                          // 先自增，保证下面除数的 n ≥ 1 / increment first so the divisor is at least one
        fDelta   := fSample - fMeanInt;                     // 新样本偏差 / deviation of the new sample
        fMeanInt := fMeanInt + (fDelta / UDINT_TO_LREAL(nAcc));     // Welford 均值递推 / Welford mean update
        fM2      := fM2 + (fDelta * (fSample - fMeanInt));          // Welford 二阶矩递推 / Welford second moment update
    END_IF
END_IF

// 段 5｜阶段机与出口发布：ENUM + CASE + ELSE 兜底，每分支内不留跨拍中间量 / segment 5, the stage machine
CASE eStage OF
    eWelfordIdle, eWelfordAccum:
        fMean  := fMeanInt;                         // 空相时内部均值恒 0，两相共用一条发布路径 / the internal mean is zero when empty, so both stages share one path
        fVar   := DL_ZERO_L;                        // 不足两样本，方差按契约置 0 / fewer than two samples, the variance is zero by contract
        fStd   := DL_ZERO_L;                        // 标准差同步置 0 / the deviation is zero as well
        bValid := FALSE;                            // 三件套不可用 / the outputs are unusable
        IF nAcc >= DL_TWO THEN
            eStage := eWelfordReady;                // 进入可用相 / enter the ready stage
        ELSIF nAcc = 0 THEN
            eStage := eWelfordIdle;                 // 回落空闲相（复位后）/ fall back to idle after a reset
        ELSE
            eStage := eWelfordAccum;                // 停在单样本相 / stay at the single sample stage
        END_IF
    eWelfordReady:
        fMean := fMeanInt;                          // 均值 / the mean
        IF nAcc > DL_ONE THEN
            fVarInt := fM2 / UDINT_TO_LREAL(nAcc - DL_ONE);     // 样本方差，分母 n−1 / sample variance
        ELSE
            fVarInt := DL_ZERO_L;                   // 结构性不可达，兜底防除零 / unreachable guard against a zero divisor
        END_IF
        IF fVarInt < DL_ZERO_L THEN
            fVarInt := DL_ZERO_L;                   // 数值负偏兜底，方差不得为负 / a numeric undershoot must not go negative
        END_IF
        fVar   := fVarInt;                          // 出口方差 / publish the variance
        fStd   := SQRT(fVarInt);                    // 出口标准差 / publish the deviation
        bValid := TRUE;                             // 三件套可用 / every output is usable
        IF nAcc < DL_TWO THEN
            IF nAcc = 0 THEN
                eStage := eWelfordIdle;             // 复位后回落空闲相 / fall back after a reset
            ELSE
                eStage := eWelfordAccum;            // 回落单样本相 / fall back to the single sample stage
            END_IF
        END_IF
ELSE
    eStage := eWelfordIdle;                         // 非法阶段拦截并复位 / intercept an illegal stage and recover
    fMean  := DL_ZERO_L;
    fVar   := DL_ZERO_L;
    fStd   := DL_ZERO_L;
    bValid := FALSE;
END_CASE

// 段 6｜计数出口：与阶段机解耦，无条件映射 / segment 6, publish the count independently of the stage machine
nCount := nAcc;                                     // 已纳入样本数 / accepted sample count
END_FUNCTION_BLOCK
